  MoveL 742 to (62.2, -35.66, 5.28) mm, rotated rx 90 ry -59.82 rz 90 deg; joints [18.012, -65.128, 129.561, -160.179, 65.77, 111.765]
  MoveL 743 to (62.59, -36.33, 5.7) mm, rotated rx 90 ry -55.77 rz 90 deg; joints [17.262, -66.589, 129.722, -160.795, 64.433, 115.685]
  MoveL 744 to (62.99, -36.97, 6.17) mm, rotated rx 90 ry -51.71 rz 90 deg; joints [16.443, -67.973, 129.873, -161.501, 63.144, 119.692]
  MoveL 745 to (63.38, -37.58, 6.68) mm, rotated rx 90 ry -47.66 rz 90 deg; joints [15.557, -69.273, 130.015, -162.302, 61.911, 123.796]
  MoveL 746 to (63.82, -38.19, 7.29) mm, rotated rx 90 ry -43.28 rz 90 deg; joints [14.528, -70.576, 130.159, -163.275, 60.653, 128.346]
  MoveL 747 to (64.25, -38.76, 7.94) mm, rotated rx 90 ry -38.89 rz 90 deg; joints [13.429, -71.764, 130.295, -164.361, 59.485, 133.017]
  MoveL 748 to (64.69, -39.27, 8.63) mm, rotated rx 90 ry -34.51 rz 90 deg; joints [12.267, -72.829, 130.424, -165.558, 58.421, 137.808]
  MoveL 749 to (65.12, -39.73, 9.35) mm, rotated rx 90 ry -30.13 rz 90 deg; joints [11.047, -73.766, 130.549, -166.865, 57.475, 142.721]
  MoveL 750 to (65.56, -40.15, 10.14) mm, rotated rx 90 ry -25.6 rz 90 deg; joints [9.732, -74.593, 130.674, -168.322, 56.634, 147.917]
  MoveL 751 to (66, -40.5, 10.96) mm, rotated rx 90 ry -21.07 rz 90 deg; joints [8.373, -75.268, 130.796, -169.878, 55.946, 153.223]
  MoveL 752 to (66.44, -40.78, 11.8) mm, rotated rx 90 ry -16.54 rz 90 deg; joints [6.977, -75.787, 130.915, -171.517, 55.423, 158.623]
  MoveL 753 to (66.88, -41, 12.66) mm, rotated rx 90 ry -12.01 rz 90 deg; joints [5.554, -76.145, 131.032, -173.221, 55.076, 164.098]
  MoveL 754 to (67.32, -41.15, 13.54) mm, rotated rx 90 ry -7.48 rz 90 deg; joints [4.115, -76.339, 131.148, -174.969, 54.913, 169.623]
  MoveL 755 to (67.76, -41.23, 14.42) mm, rotated rx 90 ry -2.95 rz 90 deg; joints [2.671, -76.366, 131.26, -176.737, 54.937, 175.174]
  MoveL 756 to (68.16, -41.25, 15.26) mm, rotated rx 90 ry 0 rz 90 deg; joints [1.719, -76.288, 131.323, -177.903, 55.053, 178.798]
  MoveL 757 to (68.57, -41.25, 16.1) mm, rotated rx 90 ry 0 rz 90 deg; joints [1.676, -76.267, 131.295, -177.955, 55.045, 178.828]
  MoveL 758 to (68.97, -41.25, 16.94) mm, rotated rx 90 ry 0 rz 90 deg; joints [1.634, -76.246, 131.266, -178.007, 55.037, 178.857]
  MoveL 759 to (69.37, -41.25, 17.77) mm, rotated rx 90 ry 0 rz 90 deg; joints [1.591, -76.225, 131.238, -178.058, 55.028, 178.887]
  MoveL 760 to (69.78, -41.25, 18.61) mm, rotated rx 90 ry 0 rz 90 deg; joints [1.548, -76.204, 131.209, -178.11, 55.02, 178.916]
  MoveL 761 to (70.18, -41.25, 19.45) mm, rotated rx 90 ry 0 rz 90 deg; joints [1.506, -76.182, 131.181, -178.162, 55.012, 178.946]
  MoveL 762 to (72.7, -41.25, 24.26) mm, rotated rx 90 ry 0 rz 90 deg; joints [1.262, -76.049, 131.001, -178.459, 54.962, 179.115]
  MoveL 763 to (75.1, -41.25, 27.7) mm, rotated rx 90 ry 0 rz 90 deg; joints [1.087, -75.919, 130.826, -178.671, 54.914, 179.236]
  MoveL 764 to (78.13, -41.25, 30.71) mm, rotated rx 90 ry 0 rz 90 deg; joints [0.934, -75.754, 130.602, -178.857, 54.854, 179.342]
  MoveL 765 to (81.19, -41.25, 33.72) mm, rotated rx 90 ry 0 rz 90 deg; joints [0.782, -75.586, 130.375, -179.042, 54.793, 179.448]
  MoveL 766 to (82.71, -41.25, 36.56) mm, rotated rx 90 ry 0 rz 90 deg; joints [0.64, -75.504, 130.263, -179.216, 54.762, 179.548]
  MoveL 767 to (83.13, -41.25, 40.01) mm, rotated rx 90 ry 0 rz 90 deg; joints [0.469, -75.482, 130.234, -179.426, 54.753, 179.669]
  MoveL 768 to (82.53, -41.25, 43.6) mm, rotated rx 90 ry 0 rz 90 deg; joints [0.291, -75.517, 130.281, -179.644, 54.765, 179.795]
  MoveL 769 to (82.18, -41.25, 44.44) mm, rotated rx 90 ry 0 rz 90 deg; joints [0.25, -75.537, 130.308, -179.694, 54.772, 179.824]
  MoveL 770 to (81.83, -41.25, 45.27) mm, rotated rx 90 ry 1.37 rz 90 deg; joints [-0.208, -75.494, 130.36, 179.746, 54.866, -178.482]
  MoveL 771 to (81.47, -41.2, 46.1) mm, rotated rx 90 ry 5.62 rz 90 deg; joints [-1.527, -75.226, 130.461, 178.141, 55.25, -173.325]
  MoveL 772 to (80.96, -41.11, 46.79) mm, rotated rx 90 ry 9.15 rz 90 deg; joints [-2.612, -74.904, 130.558, 176.838, 55.695, -169.062]
  MoveL 773 to (80.45, -40.98, 47.47) mm, rotated rx 90 ry 12.69 rz 90 deg; joints [-3.676, -74.483, 130.651, 175.577, 56.246, -164.844]
  MoveL 774 to (79.95, -40.8, 48.15) mm, rotated rx 90 ry 16.23 rz 90 deg; joints [-4.716, -73.965, 130.737, 174.367, 56.9, -160.682]
  MoveL 775 to (78.97, -40.58, 48.81) mm, rotated rx 90 ry 19.82 rz 90 deg; joints [-5.743, -73.366, 130.853, 173.198, 57.67, -156.527]
  MoveL 776 to (78, -40.32, 49.47) mm, rotated rx 90 ry 23.41 rz 90 deg; joints [-6.737, -72.67, 130.961, 172.095, 58.534, -152.445]
  MoveL 777 to (77.24, -40.22, 49.7) mm, rotated rx 90 ry 24.7 rz 90 deg; joints [-7.087, -72.418, 131.028, 171.713, 58.876, -150.995]
  MoveL 778 to (76.48, -40.11, 49.93) mm, rotated rx 90 ry 25.99 rz 90 deg; joints [-7.433, -72.154, 131.094, 171.34, 59.229, -149.556]
  MoveL 779 to (75.72, -40, 50.16) mm, rotated rx 90 ry 27.28 rz 90 deg; joints [-7.774, -71.878, 131.159, 170.977, 59.593, -148.127]
  MoveL 780 to (74.77, -39.93, 50.28) mm, rotated rx 90 ry 27.99 rz 90 deg; joints [-7.964, -71.747, 131.234, 170.777, 59.813, -147.34]
  MoveL 781 to (73.82, -39.87, 50.4) mm, rotated rx 90 ry 28.71 rz 90 deg; joints [-8.153, -71.611, 131.309, 170.579, 60.036, -146.557]
  MoveL 782 to (72.87, -39.8, 50.53) mm, rotated rx 90 ry 29.42 rz 90 deg; joints [-8.34, -71.472, 131.384, 170.384, 60.262, -145.776]
  MoveL 783 to (71.92, -39.73, 50.65) mm, rotated rx 90 ry 30.13 rz 90 deg; joints [-8.525, -71.329, 131.457, 170.192, 60.491, -144.999]
  MoveL 784 to (70.97, -39.66, 50.77) mm, rotated rx 90 ry 30.85 rz 90 deg; joints [-8.709, -71.182, 131.531, 170.003, 60.724, -144.226]
  MoveL 785 to (70.02, -39.59, 50.89) mm, rotated rx 90 ry 31.56 rz 90 deg; joints [-8.892, -71.032, 131.604, 169.817, 60.96, -143.456]
  MoveL 786 to (69.07, -39.51, 51.01) mm, rotated rx 90 ry 32.27 rz 90 deg; joints [-9.073, -70.877, 131.676, 169.633, 61.199, -142.688]
  MoveL 787 to (68.12, -39.44, 51.12) mm, rotated rx 90 ry 32.99 rz 90 deg; joints [-9.252, -70.719, 131.748, 169.452, 61.441, -141.924]
  MoveL 788 to (67.17, -39.36, 51.24) mm, rotated rx 90 ry 33.7 rz 90 deg; joints [-9.43, -70.557, 131.819, 169.274, 61.686, -141.163]
  MoveL 789 to (66.22, -39.32, 51.3) mm, rotated rx 90 ry 34.04 rz 90 deg; joints [-9.518, -70.503, 131.891, 169.187, 61.817, -140.804]
  MoveL 790 to (65.27, -39.28, 51.35) mm, rotated rx 90 ry 34.38 rz 90 deg; joints [-9.606, -70.449, 131.962, 169.101, 61.949, -140.445]
  MoveL 791 to (64.32, -39.25, 51.41) mm, rotated rx 90 ry 34.72 rz 90 deg; joints [-9.693, -70.393, 132.034, 169.015, 62.081, -140.087]
  MoveL 792 to (63.37, -39.21, 51.46) mm, rotated rx 90 ry 35.06 rz 90 deg; joints [-9.78, -70.337, 132.105, 168.93, 62.215, -139.73]
  MoveL 793 to (62.41, -39.17, 51.52) mm, rotated rx 90 ry 35.4 rz 90 deg; joints [-9.866, -70.279, 132.176, 168.846, 62.348, -139.375]
  MoveL 794 to (61.46, -39.13, 51.57) mm, rotated rx 90 ry 35.74 rz 90 deg; joints [-9.953, -70.221, 132.247, 168.762, 62.483, -139.019]
  MoveL 795 to (60.51, -39.09, 51.62) mm, rotated rx 90 ry 36.08 rz 90 deg; joints [-10.039, -70.162, 132.318, 168.679, 62.619, -138.664]
  MoveL 796 to (59.55, -39.05, 51.68) mm, rotated rx 90 ry 36.41 rz 90 deg; joints [-10.124, -70.101, 132.388, 168.596, 62.755, -138.31]
  MoveL 797 to (58.6, -39.01, 51.73) mm, rotated rx 90 ry 36.75 rz 90 deg; joints [-10.21, -70.04, 132.459, 168.514, 62.892, -137.957]
  MoveL 798 to (57.65, -39.01, 51.73) mm, rotated rx 90 ry 36.77 rz 90 deg; joints [-10.223, -70.079, 132.531, 168.503, 62.925, -137.938]
  MoveL 799 to (56.69, -39.01, 51.74) mm, rotated rx 90 ry 36.79 rz 90 deg; joints [-10.236, -70.119, 132.603, 168.491, 62.958, -137.917]
  MoveL 800 to (55.73, -39.01, 51.74) mm, rotated rx 90 ry 36.81 rz 90 deg; joints [-10.249, -70.158, 132.674, 168.48, 62.991, -137.898]
  MoveL 801 to (54.78, -39, 51.74) mm, rotated rx 90 ry 36.83 rz 90 deg; joints [-10.262, -70.198, 132.746, 168.469, 63.024, -137.878]
  MoveL 802 to (53.82, -39, 51.75) mm, rotated rx 90 ry 36.85 rz 90 deg; joints [-10.275, -70.237, 132.818, 168.457, 63.057, -137.859]
  MoveL 803 to (52.87, -39, 51.75) mm, rotated rx 90 ry 36.87 rz 90 deg; joints [-10.288, -70.276, 132.89, 168.446, 63.09, -137.84]
  MoveL 804 to (51.91, -39, 51.75) mm, rotated rx 90 ry 36.9 rz 90 deg; joints [-10.302, -70.316, 132.962, 168.435, 63.123, -137.819]
  MoveL 805 to (50.96, -38.99, 51.76) mm, rotated rx 90 ry 36.91 rz 90 deg; joints [-10.315, -70.355, 133.033, 168.423, 63.156, -137.8]
  MoveL 806 to (50, -38.99, 51.76) mm, rotated rx 90 ry 36.94 rz 90 deg; joints [-10.328, -70.394, 133.105, 168.412, 63.189, -137.781]
  MoveL 807 to (50, -39.55, 50.95) mm, rotated rx 90 ry 31.94 rz 90 deg; joints [-9.143, -71.919, 133.112, 169.592, 61.592, -143.063]
  MoveL 808 to (50, -40.03, 50.1) mm, rotated rx 90 ry 26.95 rz 90 deg; joints [-7.863, -73.276, 133.093, 170.923, 60.129, -148.499]
  MoveL 809 to (50, -40.43, 49.21) mm, rotated rx 90 ry 21.96 rz 90 deg; joints [-6.498, -74.456, 133.053, 172.398, 58.821, -154.088]
  MoveL 810 to (50, -40.76, 48.28) mm, rotated rx 90 ry 16.97 rz 90 deg; joints [-5.059, -75.448, 132.995, 174.011, 57.688, -159.823]
  MoveL 811 to (50, -41.01, 47.33) mm, rotated rx 90 ry 11.98 rz 90 deg; joints [-3.556, -76.246, 132.923, 175.747, 56.75, -165.689]
  MoveL 812 to (50, -41.17, 46.37) mm, rotated rx 90 ry 6.98 rz 90 deg; joints [-2.003, -76.843, 132.841, 177.585, 56.022, -171.665]
  MoveL 813 to (50, -41.24, 45.39) mm, rotated rx 90 ry 1.99 rz 90 deg; joints [-0.413, -77.235, 132.752, 179.499, 55.517, -177.724]
  MoveL 814 to (50, -41.25, 44.41) mm, rotated rx 90 ry 0 rz 90 deg; joints [0.258, -77.334, 132.714, -179.686, 55.381, 179.822]
  MoveL 815 to (45.62, -41.25, 43.91) mm, rotated rx 90 ry 0 rz 90 deg; joints [0.285, -77.581, 133.039, -179.654, 55.459, 179.804]
  MoveL 816 to (41.42, -41.25, 43.16) mm, rotated rx 90 ry 0 rz 90 deg; joints [0.325, -77.817, 133.349, -179.606, 55.532, 179.777]
  MoveL 817 to (38.6, -41.25, 42.58) mm, rotated rx 90 ry 0 rz 90 deg; joints [0.355, -77.977, 133.557, -179.57, 55.581, 179.757]
  MoveL 818 to (35.9, -41.25, 41.66) mm, rotated rx 90 ry 0 rz 90 deg; joints [0.404, -78.13, 133.756, -179.511, 55.627, 179.724]
  MoveL 819 to (34.18, -41.25, 39.31) mm, rotated rx 90 ry 0 rz 90 deg; joints [0.526, -78.226, 133.881, -179.363, 55.657, 179.641]
  MoveL 820 to (33.35, -41.25, 35.37) mm, rotated rx 90 ry 0 rz 90 deg; joints [0.731, -78.271, 133.939, -179.115, 55.672, 179.501]
  MoveL 821 to (33.65, -41.25, 31.56) mm, rotated rx 90 ry 0 rz 90 deg; joints [0.928, -78.25, 133.913, -178.876, 55.668, 179.366]
  MoveL 822 to (34.41, -41.25, 27.86) mm, rotated rx 90 ry 0 rz 90 deg; joints [1.119, -78.203, 133.852, -178.645, 55.656, 179.235]
  MoveL 823 to (35.45, -41.25, 23.18) mm, rotated rx 90 ry 0 rz 90 deg; joints [1.36, -78.139, 133.768, -178.352, 55.64, 179.07]
  MoveL 824 to (36.64, -41.25, 18.45) mm, rotated rx 90 ry 0 rz 90 deg; joints [1.603, -78.064, 133.671, -178.057, 55.622, 178.903]
  MoveL 825 to (36.94, -41.25, 17.47) mm, rotated rx 90 ry 0 rz 90 deg; joints [1.653, -78.046, 133.647, -177.997, 55.618, 178.868]
  MoveL 826 to (37.24, -41.25, 16.5) mm, rotated rx 90 ry 0 rz 90 deg; joints [1.703, -78.027, 133.623, -177.936, 55.613, 178.834]
  MoveL 827 to (37.53, -41.25, 15.52) mm, rotated rx 90 ry 0 rz 90 deg; joints [1.753, -78.009, 133.599, -177.876, 55.608, 178.8]
  MoveL 828 to (37.83, -41.24, 14.55) mm, rotated rx 90 ry -2.31 rz 90 deg; joints [2.533, -78.043, 133.502, -176.925, 55.498, 175.947]
  MoveL 829 to (38.13, -41.16, 13.57) mm, rotated rx 90 ry -7.28 rz 90 deg; joints [4.156, -77.984, 133.319, -174.951, 55.439, 169.855]
  MoveL 830 to (38.43, -41.02, 12.72) mm, rotated rx 90 ry -11.71 rz 90 deg; joints [5.597, -77.754, 133.151, -173.21, 55.585, 164.443]
  MoveL 831 to (38.73, -40.81, 11.87) mm, rotated rx 90 ry -16.14 rz 90 deg; joints [7.021, -77.363, 132.981, -171.512, 55.912, 159.081]
  MoveL 832 to (39.03, -40.53, 11.05) mm, rotated rx 90 ry -20.57 rz 90 deg; joints [8.417, -76.813, 132.81, -169.88, 56.412, 153.793]
  MoveL 833 to (39.33, -40.2, 10.25) mm, rotated rx 90 ry -25 rz 90 deg; joints [9.777, -76.11, 132.637, -168.329, 57.076, 148.595]
  MoveL 834 to (39.63, -39.8, 9.47) mm, rotated rx 90 ry -29.43 rz 90 deg; joints [11.09, -75.258, 132.461, -166.874, 57.89, 143.505]
  MoveL 835 to (40, -39.28, 8.64) mm, rotated rx 90 ry -34.42 rz 90 deg; joints [12.506, -74.128, 132.257, -165.363, 58.971, 137.91]
  MoveL 836 to (40.37, -38.69, 7.86) mm, rotated rx 90 ry -39.41 rz 90 deg; joints [13.843, -72.827, 132.045, -163.996, 60.205, 132.475]
  MoveL 837 to (40.74, -38.04, 7.13) mm, rotated rx 90 ry -44.41 rz 90 deg; joints [15.092, -71.368, 131.825, -162.778, 61.571, 127.199]
  MoveL 838 to (41.11, -37.32, 6.46) mm, rotated rx 90 ry -49.4 rz 90 deg; joints [16.246, -69.763, 131.594, -161.709, 63.05, 122.081]
  MoveL 839 to (41.48, -36.55, 5.85) mm, rotated rx 90 ry -54.41 rz 90 deg; joints [17.302, -68.016, 131.349, -160.783, 64.628, 117.092]
  MoveL 840 to (41.84, -35.72, 5.31) mm, rotated rx 90 ry -59.43 rz 90 deg; joints [18.249, -66.15, 131.09, -159.998, 66.28, 112.244]
  MoveL 841 to (42.21, -34.85, 4.85) mm, rotated rx 90 ry -64.44 rz 90 deg; joints [19.084, -64.176, 130.813, -159.35, 67.99, 107.521]
  MoveL 842 to (42.58, -33.95, 4.47) mm, rotated rx 90 ry -69.45 rz 90 deg; joints [19.803, -62.112, 130.519, -158.83, 69.742, 102.91]
  MoveL 843 to (42.94, -33.17, 4.21) mm, rotated rx 90 ry -73.65 rz 90 deg; joints [20.313, -60.322, 130.255, -158.491, 71.229, 99.121]
  MoveL 844 to (43.3, -32.37, 4) mm, rotated rx 90 ry -77.85 rz 90 deg; joints [20.739, -58.488, 129.978, -158.233, 72.728, 95.387]
  MoveL 845 to (43.66, -31.56, 3.86) mm, rotated rx 90 ry -82.05 rz 90 deg; joints [21.079, -56.619, 129.687, -158.055, 74.232, 91.701]
  MoveL 846 to (44.02, -30.74, 3.77) mm, rotated rx 90 ry -86.25 rz 90 deg; joints [21.333, -54.723, 129.384, -157.953, 75.735, 88.05]
  MoveL 847 to (44.51, -29.87, 3.75) mm, rotated rx 0 ry -90 rz 180 deg; joints [21.484, -53.003, 129.092, -157.928, 77.072, 84.817]
  MoveL 848 to (44.99, -29, 3.75) mm, rotated rx 0 ry -90 rz 180 deg; joints [21.476, -52.928, 129.05, -157.94, 77.102, 84.831]
  MoveL 849 to (45.47, -28.14, 3.75) mm, rotated rx 0 ry -90 rz 180 deg; joints [21.467, -52.853, 129.007, -157.951, 77.132, 84.846]
  MoveL 850 to (45.95, -27.27, 3.75) mm, rotated rx 0 ry -90 rz 180 deg; joints [21.459, -52.778, 128.965, -157.963, 77.162, 84.861]
  MoveL 851 to (47.84, -24.64, 3.75) mm, rotated rx 0 ry -90 rz 180 deg; joints [21.426, -52.538, 128.807, -158.003, 77.234, 84.899]
  MoveL 852 to (48.85, -23.61, 3.75) mm, rotated rx 0 ry -90 rz 180 deg; joints [21.408, -52.437, 128.724, -158.023, 77.25, 84.91]
  MoveL 853 to (50, -22.99, 3.75) mm, rotated rx 0 ry -90 rz 180 deg; joints [21.388, -52.36, 128.634, -158.042, 77.236, 84.91]
  MoveL 854 to (51.15, -23.61, 3.75) mm, rotated rx 0 ry -90 rz 180 deg; joints [21.368, -52.37, 128.555, -158.055, 77.151, 84.88]
  MoveL 855 to (52.16, -24.64, 3.75) mm, rotated rx 0 ry -90 rz 180 deg; joints [21.351, -52.413, 128.489, -158.063, 77.049, 84.842]
  MoveL 856 to (54.05, -27.27, 3.75) mm, rotated rx 0 ry -90 rz 180 deg; joints [21.318, -52.542, 128.371, -158.075, 76.817, 84.755]
  MoveL 857 to (54.53, -28.14, 3.75) mm, rotated rx 0 ry -90 rz 180 deg; joints [21.31, -52.589, 128.343, -158.077, 76.747, 84.728]
  MoveL 858 to (55.01, -29, 3.75) mm, rotated rx 0 ry -90 rz 180 deg; joints [21.302, -52.635, 128.314, -158.079, 76.676, 84.701]
  MoveL 859 to (55.49, -29.87, 3.75) mm, rotated rx 0 ry -90 rz 180 deg; joints [21.293, -52.681, 128.285, -158.081, 76.606, 84.675]
  MoveL 860 to (55.98, -30.74, 3.77) mm, rotated rx 90 ry -86.25 rz 90 deg; joints [21.127, -54.352, 128.505, -158.116, 75.243, 87.907]
  MoveL 861 to (56.34, -31.56, 3.86) mm, rotated rx 90 ry -82.05 rz 90 deg; joints [20.863, -56.201, 128.753, -158.223, 73.729, 91.562]
  MoveL 862 to (56.7, -32.37, 4) mm, rotated rx 90 ry -77.85 rz 90 deg; joints [20.513, -58.02, 128.989, -158.407, 72.217, 95.256]
  MoveL 863 to (57.06, -33.17, 4.21) mm, rotated rx 90 ry -73.65 rz 90 deg; joints [20.08, -59.803, 129.212, -158.67, 70.712, 98.998]
  MoveL 864 to (57.42, -33.95, 4.47) mm, rotated rx 90 ry -69.45 rz 90 deg; joints [19.563, -61.538, 129.422, -159.014, 69.221, 102.798]
  MoveL 865 to (57.79, -34.85, 4.85) mm, rotated rx 90 ry -64.44 rz 90 deg; joints [18.84, -63.54, 129.66, -159.537, 67.472, 107.424]
  MoveL 866 to (58.16, -35.72, 5.31) mm, rotated rx 90 ry -59.43 rz 90 deg; joints [18.003, -65.448, 129.881, -160.188, 65.768, 112.163]
  MoveL 867 to (58.52, -36.55, 5.85) mm, rotated rx 90 ry -54.41 rz 90 deg; joints [17.056, -67.249, 130.086, -160.974, 64.123, 117.028]
  MoveL 868 to (58.89, -37.32, 6.46) mm, rotated rx 90 ry -49.4 rz 90 deg; joints [16.003, -68.928, 130.277, -161.901, 62.555, 122.035]
  MoveL 869 to (59.26, -38.04, 7.13) mm, rotated rx 90 ry -44.41 rz 90 deg; joints [14.856, -70.466, 130.453, -162.969, 61.088, 127.169]
  MoveL 870 to (59.63, -38.69, 7.86) mm, rotated rx 90 ry -39.41 rz 90 deg; joints [13.616, -71.858, 130.619, -164.183, 59.733, 132.46]
  MoveL 871 to (60, -39.28, 8.64) mm, rotated rx 90 ry -34.42 rz 90 deg; joints [12.292, -73.092, 130.777, -165.543, 58.512, 137.908]
  MoveL 872 to (60.37, -39.8, 9.47) mm, rotated rx 90 ry -29.43 rz 90 deg; joints [10.892, -74.158, 130.928, -167.045, 57.443, 143.514]
  MoveL 873 to (60.67, -40.2, 10.25) mm, rotated rx 90 ry -25 rz 90 deg; joints [9.596, -74.957, 131.059, -168.487, 56.639, 148.61]
  MoveL 874 to (60.97, -40.53, 11.05) mm, rotated rx 90 ry -20.57 rz 90 deg; joints [8.256, -75.61, 131.188, -170.023, 55.983, 153.812]
  MoveL 875 to (61.27, -40.81, 11.87) mm, rotated rx 90 ry -16.14 rz 90 deg; joints [6.883, -76.113, 131.314, -171.638, 55.488, 159.101]
  MoveL 876 to (61.57, -41.02, 12.72) mm, rotated rx 90 ry -11.71 rz 90 deg; joints [5.484, -76.46, 131.438, -173.314, 55.162, 164.462]
  MoveL 877 to (61.87, -41.16, 13.57) mm, rotated rx 90 ry -7.28 rz 90 deg; joints [4.07, -76.649, 131.561, -175.031, 55.013, 169.87]
  MoveL 878 to (62.17, -41.24, 14.55) mm, rotated rx 90 ry -2.31 rz 90 deg; joints [2.479, -76.673, 131.698, -176.976, 55.062, 175.957]
  MoveL 879 to (62.47, -41.25, 15.52) mm, rotated rx 90 ry 0 rz 90 deg; joints [1.714, -76.607, 131.749, -177.911, 55.16, 178.806]
  MoveL 880 to (62.76, -41.25, 16.5) mm, rotated rx 90 ry 0 rz 90 deg; joints [1.665, -76.592, 131.729, -177.971, 55.154, 178.841]
  MoveL 881 to (63.06, -41.25, 17.47) mm, rotated rx 90 ry 0 rz 90 deg; joints [1.615, -76.576, 131.709, -178.032, 55.148, 178.875]
  MoveL 882 to (63.36, -41.25, 18.45) mm, rotated rx 90 ry 0 rz 90 deg; joints [1.565, -76.561, 131.689, -178.092, 55.142, 178.909]
  MoveL 883 to (64.55, -41.25, 23.18) mm, rotated rx 90 ry 0 rz 90 deg; joints [1.325, -76.501, 131.609, -178.384, 55.118, 179.076]
  MoveL 884 to (65.59, -41.25, 27.86) mm, rotated rx 90 ry 0 rz 90 deg; joints [1.088, -76.449, 131.539, -178.673, 55.097, 179.241]
  MoveL 885 to (66.35, -41.25, 31.56) mm, rotated rx 90 ry 0 rz 90 deg; joints [0.901, -76.41, 131.486, -178.901, 55.081, 179.371]
  MoveL 886 to (66.65, -41.25, 35.37) mm, rotated rx 90 ry 0 rz 90 deg; joints [0.709, -76.396, 131.468, -179.135, 55.075, 179.505]
  MoveL 887 to (65.82, -41.25, 39.31) mm, rotated rx 90 ry 0 rz 90 deg; joints [0.511, -76.445, 131.533, -179.376, 55.09, 179.643]
  MoveL 888 to (64.11, -41.25, 41.66) mm, rotated rx 90 ry 0 rz 90 deg; joints [0.394, -76.542, 131.663, -179.52, 55.122, 179.726]
  MoveL 889 to (61.4, -41.25, 42.58) mm, rotated rx 90 ry 0 rz 90 deg; joints [0.348, -76.693, 131.865, -179.576, 55.172, 179.758]
  MoveL 890 to (58.58, -41.25, 43.16) mm, rotated rx 90 ry 0 rz 90 deg; joints [0.32, -76.852, 132.075, -179.611, 55.225, 179.778]
  MoveL 891 to (54.38, -41.25, 43.91) mm, rotated rx 90 ry 0 rz 90 deg; joints [0.283, -77.087, 132.388, -179.656, 55.301, 179.804]
  MoveL 892 to (50, -41.25, 44.41) mm, rotated rx 90 ry 0 rz 90 deg; joints [0.258, -77.334, 132.714, -179.686, 55.381, 179.822]
  MoveL 893 to (50, -41.25, 34.01) mm, rotated rx 90 ry 0 rz 90 deg; joints [0.789, -77.328, 132.707, -179.041, 55.382, 179.455]
  MoveL 894 to (47.54, -41.25, 33.12) mm, rotated rx 90 ry 0 rz 90 deg; joints [0.837, -77.466, 132.888, -178.984, 55.426, 179.423]
  MoveL 895 to (45.56, -41.25, 31.05) mm, rotated rx 90 ry 0 rz 90 deg; joints [0.944, -77.576, 133.033, -178.854, 55.462, 179.35]
  MoveL 896 to (44.02, -41.25, 28.52) mm, rotated rx 90 ry 0 rz 90 deg; joints [1.075, -77.661, 133.144, -178.695, 55.49, 179.261]
  MoveL 897 to (42.9, -41.25, 25.95) mm, rotated rx 90 ry 0 rz 90 deg; joints [1.209, -77.721, 133.223, -178.534, 55.511, 179.17]
  MoveL 898 to (41.78, -41.25, 20.71) mm, rotated rx 90 ry 0 rz 90 deg; joints [1.479, -77.777, 133.297, -178.205, 55.532, 178.984]
  MoveL 899 to (41.91, -41.25, 15.28) mm, rotated rx 90 ry 0 rz 90 deg; joints [1.758, -77.761, 133.275, -177.867, 55.533, 178.792]
  MoveL 900 to (42.06, -41.23, 14.35) mm, rotated rx 90 ry -3.31 rz 90 deg; joints [2.851, -77.812, 133.158, -176.535, 55.395, 174.716]
  MoveL 901 to (42.21, -41.14, 13.42) mm, rotated rx 90 ry -8.05 rz 90 deg; joints [4.394, -77.728, 132.993, -174.659, 55.381, 168.907]
  MoveL 902 to (42.36, -40.97, 12.51) mm, rotated rx 90 ry -12.79 rz 90 deg; joints [5.926, -77.458, 132.826, -172.81, 55.579, 163.133]
  MoveL 903 to (42.51, -40.73, 11.61) mm, rotated rx 90 ry -17.52 rz 90 deg; joints [7.437, -77.003, 132.657, -171.016, 55.982, 157.42]
  MoveL 904 to (42.72, -40.43, 10.78) mm, rotated rx 90 ry -22.06 rz 90 deg; joints [8.851, -76.397, 132.488, -169.373, 56.549, 152.035]
  MoveL 905 to (42.93, -40.06, 9.96) mm, rotated rx 90 ry -26.6 rz 90 deg; joints [10.225, -75.632, 132.318, -167.82, 57.282, 146.75]
  MoveL 906 to (43.13, -39.63, 9.18) mm, rotated rx 90 ry -31.13 rz 90 deg; joints [11.547, -74.714, 132.144, -166.372, 58.167, 141.581]
  MoveL 907 to (43.34, -39.14, 8.44) mm, rotated rx 90 ry -35.67 rz 90 deg; joints [12.811, -73.651, 131.965, -165.039, 59.19, 136.539]
  MoveL 908 to (43.6, -38.61, 7.76) mm, rotated rx 90 ry -40.05 rz 90 deg; joints [13.968, -72.49, 131.783, -163.865, 60.294, 131.794]
  MoveL 909 to (43.86, -38.03, 7.12) mm, rotated rx 90 ry -44.43 rz 90 deg; joints [15.057, -71.209, 131.594, -162.806, 61.497, 127.171]
  MoveL 910 to (44.12, -37.41, 6.53) mm, rotated rx 90 ry -48.81 rz 90 deg; joints [16.073, -69.815, 131.397, -161.861, 62.786, 122.671]
  MoveL 911 to (44.38, -36.74, 5.99) mm, rotated rx 90 ry -53.19 rz 90 deg; joints [17.011, -68.318, 131.19, -161.029, 64.149, 118.286]
  MoveL 912 to (44.68, -36.11, 5.55) mm, rotated rx 90 ry -57.11 rz 90 deg; joints [17.78, -66.894, 130.99, -160.379, 65.418, 114.453]
  MoveL 913 to (44.99, -35.45, 5.16) mm, rotated rx 90 ry -61.03 rz 90 deg; joints [18.482, -65.401, 130.78, -159.812, 66.726, 110.702]
  MoveL 914 to (45.3, -34.76, 4.81) mm, rotated rx 90 ry -64.95 rz 90 deg; joints [19.115, -63.846, 130.559, -159.328, 68.067, 107.025]
  MoveL 915 to (45.7, -34.02, 4.49) mm, rotated rx 90 ry -69.07 rz 90 deg; joints [19.701, -62.151, 130.31, -158.905, 69.498, 103.234]
  MoveL 916 to (46.1, -33.25, 4.23) mm, rotated rx 90 ry -73.19 rz 90 deg; joints [20.208, -60.404, 130.049, -158.565, 70.948, 99.508]
  MoveL 917 to (46.5, -32.47, 4.03) mm, rotated rx 90 ry -77.31 rz 90 deg; joints [20.634, -58.615, 129.776, -158.304, 72.41, 95.837]
  MoveL 918 to (47.02, -31.63, 3.87) mm, rotated rx 90 ry -81.68 rz 90 deg; joints [20.994, -56.674, 129.464, -158.113, 73.964, 91.991]
  MoveL 919 to (47.54, -30.77, 3.78) mm, rotated rx 90 ry -86.05 rz 90 deg; joints [21.262, -54.706, 129.14, -158.005, 75.517, 88.185]
  MoveL 920 to (48.06, -29.92, 3.75) mm, rotated rx 0 ry -90 rz 180 deg; joints [21.422, -52.903, 128.832, -157.978, 76.919, 84.769]
  MoveL 921 to (49.06, -28.63, 3.75) mm, rotated rx 0 ry -90 rz 180 deg; joints [21.405, -52.783, 128.748, -157.999, 76.951, 84.787]
  MoveL 922 to (50, -27.82, 3.75) mm, rotated rx 0 ry -90 rz 180 deg; joints [21.388, -52.699, 128.673, -158.016, 76.958, 84.795]
  MoveL 923 to (50.94, -28.63, 3.75) mm, rotated rx 0 ry -90 rz 180 deg; joints [21.372, -52.729, 128.61, -158.025, 76.871, 84.763]
  MoveL 924 to (51.94, -29.92, 3.75) mm, rotated rx 0 ry -90 rz 180 deg; joints [21.355, -52.789, 128.546, -158.032, 76.754, 84.719]
  MoveL 925 to (52.46, -30.77, 3.78) mm, rotated rx 90 ry -86.05 rz 90 deg; joints [21.177, -54.553, 128.778, -158.072, 75.315, 88.126]
  MoveL 926 to (52.98, -31.63, 3.87) mm, rotated rx 90 ry -81.68 rz 90 deg; joints [20.892, -56.477, 129.025, -158.192, 73.729, 91.926]
  MoveL 927 to (53.5, -32.47, 4.03) mm, rotated rx 90 ry -77.31 rz 90 deg; joints [20.516, -58.368, 129.258, -158.395, 72.144, 95.77]
  MoveL 928 to (53.9, -33.25, 4.23) mm, rotated rx 90 ry -73.19 rz 90 deg; joints [20.079, -60.115, 129.472, -158.664, 70.663, 99.441]
  MoveL 929 to (54.3, -34.02, 4.49) mm, rotated rx 90 ry -69.07 rz 90 deg; joints [19.562, -61.816, 129.674, -159.011, 69.197, 103.17]
  MoveL 930 to (54.7, -34.76, 4.81) mm, rotated rx 90 ry -64.95 rz 90 deg; joints [18.967, -63.463, 129.863, -159.442, 67.752, 106.965]
  MoveL 931 to (55.01, -35.45, 5.16) mm, rotated rx 90 ry -61.03 rz 90 deg; joints [18.329, -64.976, 130.037, -159.93, 66.405, 110.648]
  MoveL 932 to (55.32, -36.11, 5.55) mm, rotated rx 90 ry -57.11 rz 90 deg; joints [17.623, -66.426, 130.201, -160.5, 65.092, 114.407]
  MoveL 933 to (55.62, -36.74, 5.99) mm, rotated rx 90 ry -53.19 rz 90 deg; joints [16.851, -67.806, 130.356, -161.155, 63.821, 118.247]
  MoveL 934 to (55.88, -37.41, 6.53) mm, rotated rx 90 ry -48.81 rz 90 deg; joints [15.913, -69.261, 130.525, -161.988, 62.461, 122.641]
  MoveL 935 to (56.14, -38.03, 7.12) mm, rotated rx 90 ry -44.43 rz 90 deg; joints [14.9, -70.611, 130.684, -162.932, 61.176, 127.151]
  MoveL 936 to (56.4, -38.61, 7.76) mm, rotated rx 90 ry -40.05 rz 90 deg; joints [13.816, -71.849, 130.835, -163.99, 59.978, 131.782]
  MoveL 937 to (56.66, -39.14, 8.44) mm, rotated rx 90 ry -35.67 rz 90 deg; joints [12.665, -72.966, 130.98, -165.161, 58.88, 136.536]
  MoveL 938 to (56.87, -39.63, 9.18) mm, rotated rx 90 ry -31.13 rz 90 deg; joints [11.41, -73.991, 131.127, -166.489, 57.865, 141.585]
  MoveL 939 to (57.07, -40.06, 9.96) mm, rotated rx 90 ry -26.6 rz 90 deg; joints [10.099, -74.872, 131.271, -167.93, 56.986, 146.758]
  MoveL 940 to (57.28, -40.43, 10.78) mm, rotated rx 90 ry -22.06 rz 90 deg; joints [8.739, -75.602, 131.411, -169.473, 56.26, 152.047]
  MoveL 941 to (57.49, -40.73, 11.61) mm, rotated rx 90 ry -17.52 rz 90 deg; joints [7.34, -76.175, 131.548, -171.104, 55.697, 157.434]
  MoveL 942 to (57.64, -40.97, 12.51) mm, rotated rx 90 ry -12.79 rz 90 deg; joints [5.847, -76.604, 131.695, -172.882, 55.298, 163.146]
  MoveL 943 to (57.79, -41.14, 13.42) mm, rotated rx 90 ry -8.05 rz 90 deg; joints [4.333, -76.853, 131.839, -174.714, 55.101, 168.918]
  MoveL 944 to (57.94, -41.23, 14.35) mm, rotated rx 90 ry -3.31 rz 90 deg; joints [2.811, -76.918, 131.981, -176.572, 55.111, 174.723]
  MoveL 945 to (58.09, -41.25, 15.28) mm, rotated rx 90 ry 0 rz 90 deg; joints [1.733, -76.851, 132.075, -177.89, 55.242, 178.797]
  MoveL 946 to (58.22, -41.25, 20.71) mm, rotated rx 90 ry 0 rz 90 deg; joints [1.458, -76.852, 132.076, -178.225, 55.237, 178.988]
  MoveL 947 to (57.1, -41.25, 25.95) mm, rotated rx 90 ry 0 rz 90 deg; joints [1.193, -76.922, 132.169, -178.548, 55.256, 179.172]
  MoveL 948 to (55.98, -41.25, 28.52) mm, rotated rx 90 ry 0 rz 90 deg; joints [1.064, -76.987, 132.256, -178.705, 55.275, 179.262]
  MoveL 949 to (54.44, -41.25, 31.05) mm, rotated rx 90 ry 0 rz 90 deg; joints [0.937, -77.076, 132.374, -178.86, 55.303, 179.351]
  MoveL 950 to (52.46, -41.25, 33.12) mm, rotated rx 90 ry 0 rz 90 deg; joints [0.833, -77.19, 132.524, -178.987, 55.338, 179.424]
  MoveL 951 to (50, -41.25, 34.01) mm, rotated rx 90 ry 0 rz 90 deg; joints [0.789, -77.328, 132.707, -179.041, 55.382, 179.455]
  MoveL 952 to (50, -86.25, 34.01) mm, rotated rx 90 ry 0 rz 90 deg; joints [0.789, -79.797, 131.591, -178.995, 51.799, 179.379]
  Sollgeschwindigkeit (200.0 mm/s)
  MoveL 953 to (48.17, -86.25, 38.44) mm, rotated rx 90 ry 0 rz 90 deg; joints [0.564, -79.907, 131.729, -179.282, 51.824, 179.556]
  MoveL 954 to (46.35, -86.25, 42.86) mm, rotated rx 90 ry 0 rz 90 deg; joints [0.338, -80.017, 131.865, -179.57, 51.848, 179.734]
  MoveL 955 to (44.53, -85.85, 51.72) mm, rotated rx 90 ry 6.86 rz 90 deg; joints [-2.25, -79.646, 132.15, 177.165, 52.538, -171.412]
  MoveL 956 to (42.7, -82.81, 64.37) mm, rotated rx 90 ry 20.14 rz 90 deg; joints [-6.807, -77.603, 132.547, 171.703, 55.227, -155.106]
  MoveL 957 to (40.88, -76.95, 75.98) mm, rotated rx 90 ry 33.42 rz 90 deg; joints [-10.816, -74.04, 132.838, 167.409, 59.412, -140.098]
  MoveL 958 to (39.05, -68.58, 85.93) mm, rotated rx 90 ry 46.7 rz 90 deg; joints [-14.061, -69.153, 132.929, 164.401, 64.618, -126.48]
  MoveL 959 to (37.23, -58.15, 93.7) mm, rotated rx 90 ry 59.97 rz 90 deg; joints [-16.402, -63.219, 132.732, 162.556, 70.381, -114.004]
  MoveL 960 to (35.4, -46.21, 98.86) mm, rotated rx 90 ry 73.25 rz 90 deg; joints [-17.763, -56.576, 132.191, 161.7, 76.315, -102.275]
  MoveL 961 to (33.58, -33.41, 101.15) mm, rotated rx 90 ry 86.53 rz 90 deg; joints [-18.107, -49.598, 131.303, 161.714, 82.118, -90.877]
  MoveL 962 to (31.75, -26.73, 101.25) mm, rotated rx 0 ry 90 rz 0 deg; joints [-18.048, -47.549, 131.064, 161.844, 83.835, -87.983]
  MoveL 963 to (29.93, -22.3, 101.25) mm, rotated rx 0 ry 90 rz 0 deg; joints [-18.076, -47.253, 131.124, 161.827, 84.174, -88.092]
  MoveL 964 to (28.1, -17.88, 101.25) mm, rotated rx 0 ry 90 rz 0 deg; joints [-18.104, -46.956, 131.182, 161.81, 84.513, -88.2]
  MoveL 965 to (26.28, -13.45, 101.25) mm, rotated rx 0 ry 90 rz 0 deg; joints [-18.132, -46.657, 131.238, 161.792, 84.851, -88.309]
  MoveL 966 to (24.45, -9.03, 101.25) mm, rotated rx 0 ry 90 rz 0 deg; joints [-18.16, -46.356, 131.292, 161.773, 85.188, -88.418]
  MoveL 967 to (22.63, -4.6, 101.25) mm, rotated rx 0 ry 90 rz 0 deg; joints [-18.188, -46.054, 131.343, 161.754, 85.525, -88.527]
  Sollgeschwindigkeit (50.0 mm/s)
  MoveL 968 to (22.63, -4.6, 56.25) mm, rotated rx 0 ry 90 rz 0 deg; joints [-16.036, -46.315, 132.346, 163.927, 86.186, -88.902]
  MoveL 969 to (25.24, -8.42, 56.25) mm, rotated rx 0 ry 90 rz 0 deg; joints [-16, -46.561, 132.227, 163.956, 85.834, -88.803]
  MoveL 970 to (28.39, -11.75, 56.25) mm, rotated rx 0 ry 90 rz 0 deg; joints [-15.957, -46.757, 132.057, 163.992, 85.481, -88.705]
  MoveL 971 to (31.96, -14.9, 56.25) mm, rotated rx 0 ry 90 rz 0 deg; joints [-15.908, -46.928, 131.852, 164.033, 85.119, -88.605]
  MoveL 972 to (34.49, -17.04, 56.25) mm, rotated rx 0 ry 90 rz 0 deg; joints [-15.873, -47.041, 131.704, 164.061, 84.867, -88.536]
  MoveL 973 to (37.11, -19.32, 56.25) mm, rotated rx 0 ry 90 rz 0 deg; joints [-15.838, -47.162, 131.551, 164.09, 84.603, -88.464]
  MoveL 974 to (39.78, -21.76, 56.25) mm, rotated rx 0 ry 90 rz 0 deg; joints [-15.801, -47.292, 131.396, 164.119, 84.327, -88.389]
  MoveL 975 to (42.51, -24.11, 56.25) mm, rotated rx 0 ry 90 rz 0 deg; joints [-15.765, -47.413, 131.235, 164.148, 84.055, -88.315]
  MoveL 976 to (45.72, -25.96, 56.25) mm, rotated rx 0 ry 90 rz 0 deg; joints [-15.722, -47.484, 131.029, 164.183, 83.787, -88.244]
  MoveL 977 to (50, -26.64, 56.25) mm, rotated rx 0 ry 90 rz 0 deg; joints [-15.665, -47.443, 130.724, 164.233, 83.531, -88.178]
  MoveL 978 to (54.28, -25.96, 56.25) mm, rotated rx 0 ry 90 rz 0 deg; joints [-15.608, -47.298, 130.396, 164.284, 83.353, -88.135]
  MoveL 979 to (57.49, -24.11, 56.25) mm, rotated rx 0 ry 90 rz 0 deg; joints [-15.566, -47.09, 130.128, 164.324, 83.295, -88.123]
  MoveL 980 to (60.22, -21.76, 56.25) mm, rotated rx 0 ry 90 rz 0 deg; joints [-15.53, -46.856, 129.888, 164.36, 83.288, -88.126]
  MoveL 981 to (62.89, -19.32, 56.25) mm, rotated rx 0 ry 90 rz 0 deg; joints [-15.495, -46.616, 129.65, 164.395, 83.288, -88.13]
  MoveL 982 to (65.51, -17.04, 56.25) mm, rotated rx 0 ry 90 rz 0 deg; joints [-15.461, -46.39, 129.417, 164.429, 83.281, -88.133]
  MoveL 983 to (68.04, -14.9, 56.25) mm, rotated rx 0 ry 90 rz 0 deg; joints [-15.428, -46.176, 129.192, 164.462, 83.269, -88.133]
  MoveL 984 to (71.61, -11.75, 56.25) mm, rotated rx 0 ry 90 rz 0 deg; joints [-15.383, -45.867, 128.873, 164.508, 83.258, -88.136]
  MoveL 985 to (74.76, -8.42, 56.25) mm, rotated rx 0 ry 90 rz 0 deg; joints [-15.342, -45.554, 128.581, 164.549, 83.277, -88.147]
  MoveL 986 to (77.37, -4.6, 56.25) mm, rotated rx 0 ry 90 rz 0 deg; joints [-15.309, -45.218, 128.319, 164.585, 83.347, -88.17]
  MoveL 987 to (79.31, 0, 56.25) mm, rotated rx 0 ry 90 rz 0 deg; joints [-15.284, -44.839, 128.091, 164.614, 83.492, -88.213]
  MoveL 988 to (79.31, 0, 101.25) mm, rotated rx 0 ry 90 rz 0 deg; joints [-17.348, -44.556, 127.11, 162.514, 82.895, -87.768]
  END

--- program CFLines (robot KUKA KR 30 HA) ---
  BAS (#INITMOV,0)
  BAS (#VEL_PTP,100)
  BAS (#ACC_PTP,20)
  Sollgeschwindigkeit (200.0 mm/s)
  Werkzeug setzen: TOOL 0
  Referenz erstellen.: BASE 0
  $ADVANCE = 5
  $APO.CPTP = 1.000
  $APO.CDIS = 1.000
  Sollgeschwindigkeit (1000.0 mm/s)
  Frame wechseln at (1565.36, -92.38, 870.24) mm, rotated rx -90 ry 0 rz 0 deg
  Werkzeug setzen at (355.39, 32.27, 175.35) mm
  Sollgeschwindigkeit (200.0 mm/s)
  MoveL 2 to (-44.31, -80.09, -14.44) mm, rotated rx 90 ry -30.45 rz 90 deg; joints [14.986, -80.269, 119.983, -157.269, 42.006, 132.262]
  Sollgeschwindigkeit (50.0 mm/s)
  MoveL 3 to (-44.31, -41.29, 8.36) mm, rotated rx 90 ry -30.45 rz 90 deg; joints [13.945, -79.174, 121.774, -159.855, 44.406, 134.869]
  MoveL 4 to (-43.34, -41.28, 8.34) mm, rotated rx 90 ry -30.55 rz 90 deg; joints [13.96, -79.092, 121.706, -159.84, 44.423, 134.752]
  MoveL 5 to (-42.36, -41.27, 8.32) mm, rotated rx 90 ry -30.66 rz 90 deg; joints [13.975, -79.009, 121.639, -159.824, 44.441, 134.636]
  MoveL 6 to (-41.38, -41.26, 8.3) mm, rotated rx 90 ry -30.77 rz 90 deg; joints [13.99, -78.927, 121.571, -159.808, 44.458, 134.52]
  MoveL 7 to (-40.41, -41.24, 8.28) mm, rotated rx 90 ry -30.88 rz 90 deg; joints [14.005, -78.845, 121.503, -159.793, 44.475, 134.403]
  MoveL 8 to (-39.43, -41.23, 8.26) mm, rotated rx 90 ry -30.99 rz 90 deg; joints [14.019, -78.763, 121.435, -159.777, 44.492, 134.287]
  MoveL 9 to (-38.45, -41.22, 8.23) mm, rotated rx 90 ry -31.1 rz 90 deg; joints [14.034, -78.68, 121.367, -159.762, 44.51, 134.17]
  MoveL 10 to (-37.49, -41.11, 8.06) mm, rotated rx 90 ry -32 rz 90 deg; joints [14.237, -78.418, 121.326, -159.561, 44.769, 133.176]
  MoveL 11 to (-36.53, -41, 7.88) mm, rotated rx 90 ry -32.91 rz 90 deg; joints [14.437, -78.151, 121.285, -159.367, 45.032, 132.19]
  MoveL 12 to (-35.57, -40.88, 7.71) mm, rotated rx 90 ry -33.81 rz 90 deg; joints [14.633, -77.882, 121.246, -159.18, 45.298, 131.211]
  MoveL 13 to (-34.61, -40.77, 7.54) mm, rotated rx 90 ry -34.72 rz 90 deg; joints [14.826, -77.609, 121.207, -159, 45.566, 130.239]
  MoveL 14 to (-33.65, -40.65, 7.37) mm, rotated rx 90 ry -35.62 rz 90 deg; joints [15.016, -77.333, 121.169, -158.828, 45.838, 129.275]
  MoveL 15 to (-32.69, -40.53, 7.2) mm, rotated rx 90 ry -36.53 rz 90 deg; joints [15.203, -77.054, 121.132, -158.662, 46.112, 128.318]
  MoveL 16 to (-31.8, -40.31, 6.91) mm, rotated rx 90 ry -38.11 rz 90 deg; joints [15.53, -76.603, 121.127, -158.381, 46.613, 126.661]
  MoveL 17 to (-30.9, -40.08, 6.63) mm, rotated rx 90 ry -39.69 rz 90 deg; joints [15.847, -76.142, 121.124, -158.121, 47.121, 125.026]
  MoveL 18 to (-30, -39.85, 6.36) mm, rotated rx 90 ry -41.27 rz 90 deg; joints [16.154, -75.672, 121.123, -157.88, 47.638, 123.411]
  MoveL 19 to (-29.1, -39.6, 6.09) mm, rotated rx 90 ry -42.85 rz 90 deg; joints [16.451, -75.192, 121.124, -157.659, 48.161, 121.817]
  MoveL 20 to (-28.2, -39.35, 5.83) mm, rotated rx 90 ry -44.43 rz 90 deg; joints [16.737, -74.703, 121.127, -157.457, 48.692, 120.244]
  MoveL 21 to (-27.3, -39.1, 5.58) mm, rotated rx 90 ry -46.01 rz 90 deg; joints [17.012, -74.205, 121.132, -157.274, 49.229, 118.688]
  MoveL 22 to (-26.35, -38.63, 5.15) mm, rotated rx 90 ry -48.76 rz 90 deg; joints [17.473, -73.353, 121.19, -156.991, 50.188, 116.029]
  MoveL 23 to (-25.4, -38.15, 4.75) mm, rotated rx 90 ry -51.51 rz 90 deg; joints [17.901, -72.475, 121.252, -156.759, 51.164, 113.421]
  MoveL 24 to (-24.44, -37.65, 4.37) mm, rotated rx 90 ry -54.25 rz 90 deg; joints [18.296, -71.574, 121.317, -156.575, 52.154, 110.862]
  MoveL 25 to (-23.49, -37.13, 4.01) mm, rotated rx 90 ry -57 rz 90 deg; joints [18.657, -70.65, 121.386, -156.438, 53.156, 108.347]
  MoveL 26 to (-22.54, -36.6, 3.69) mm, rotated rx 90 ry -59.74 rz 90 deg; joints [18.984, -69.705, 121.456, -156.344, 54.168, 105.873]
  MoveL 27 to (-21.71, -35.91, 3.31) mm, rotated rx 90 ry -63.19 rz 90 deg; joints [19.35, -68.512, 121.573, -156.281, 55.458, 102.823]
  MoveL 28 to (-20.88, -35.2, 2.98) mm, rotated rx 90 ry -66.63 rz 90 deg; joints [19.662, -67.292, 121.692, -156.278, 56.758, 99.824]
  MoveL 29 to (-20.05, -34.47, 2.68) mm, rotated rx 90 ry -70.08 rz 90 deg; joints [19.918, -66.048, 121.81, -156.332, 58.064, 96.871]
  MoveL 30 to (-19.22, -33.72, 2.44) mm, rotated rx 90 ry -73.52 rz 90 deg; joints [20.119, -64.783, 121.926, -156.438, 59.374, 93.956]
  MoveL 31 to (-18.39, -32.96, 2.24) mm, rotated rx 90 ry -76.96 rz 90 deg; joints [20.265, -63.501, 122.04, -156.595, 60.685, 91.072]
  MoveL 32 to (-17.57, -32.18, 2.08) mm, rotated rx 90 ry -80.4 rz 90 deg; joints [20.354, -62.209, 122.151, -156.798, 61.992, 88.215]
  MoveL 33 to (-16.74, -31.41, 1.98) mm, rotated rx 90 ry -83.84 rz 90 deg; joints [20.388, -60.907, 122.258, -157.047, 63.294, 85.379]
  MoveL 34 to (-15.92, -30.62, 1.92) mm, rotated rx 90 ry -87.28 rz 90 deg; joints [20.366, -59.601, 122.36, -157.338, 64.588, 82.557]
  MoveL 35 to (-15.1, -29.83, 1.9) mm, rotated rx 0 ry -90 rz 180 deg; joints [20.307, -58.552, 122.423, -157.6, 65.606, 80.339]
  MoveL 36 to (-14.27, -29, 1.9) mm, rotated rx 0 ry -90 rz 180 deg; joints [20.294, -58.47, 122.364, -157.618, 65.624, 80.354]
  MoveL 37 to (-12.9, -27.3, 1.9) mm, rotated rx 0 ry -90 rz 180 deg; joints [20.273, -58.315, 122.266, -157.651, 65.674, 80.388]
  MoveL 38 to (-12.11, -25.32, 1.9) mm, rotated rx 0 ry -90 rz 180 deg; joints [20.261, -58.166, 122.214, -157.68, 65.761, 80.433]
  MoveL 39 to (-12.03, -23.12, 1.9) mm, rotated rx 0 ry -90 rz 180 deg; joints [20.259, -58.033, 122.217, -157.705, 65.887, 80.49]
  MoveL 40 to (-12.95, -19.92, 1.9) mm, rotated rx 0 ry -90 rz 180 deg; joints [20.274, -57.881, 122.3, -157.729, 66.107, 80.582]
  MoveL 41 to (-14.74, -17.2, 1.9) mm, rotated rx 0 ry -90 rz 180 deg; joints [20.301, -57.791, 122.448, -157.739, 66.331, 80.668]
  MoveL 42 to (-18.88, -13.11, 1.9) mm, rotated rx 0 ry -90 rz 180 deg; joints [20.366, -57.71, 122.779, -157.738, 66.724, 80.811]
  MoveL 43 to (-23.52, -9.64, 1.9) mm, rotated rx 0 ry -90 rz 180 deg; joints [20.438, -57.683, 123.144, -157.724, 67.098, 80.942]
  MoveL 44 to (-28.63, -7.16, 1.9) mm, rotated rx 0 ry -90 rz 180 deg; joints [20.518, -57.73, 123.541, -157.693, 67.433, 81.053]
  MoveL 45 to (-33.91, -5.84, 1.9) mm, rotated rx 0 ry -90 rz 180 deg; joints [20.602, -57.854, 123.946, -157.648, 67.707, 81.134]
  MoveL 46 to (-39.38, -5.04, 1.9) mm, rotated rx 0 ry -90 rz 180 deg; joints [20.689, -58.015, 124.364, -157.594, 67.957, 81.204]
  MoveL 47 to (-44.82, -4.13, 1.9) mm, rotated rx 0 ry -90 rz 180 deg; joints [20.777, -58.168, 124.778, -157.541, 68.213, 81.277]
  MoveL 48 to (-50, -2.49, 1.9) mm, rotated rx 0 ry -90 rz 180 deg; joints [20.861, -58.263, 125.173, -157.497, 68.502, 81.367]
  MoveL 49 to (-20.13, 0, 1.9) mm, rotated rx 0 ry -90 rz 180 deg; joints [20.385, -56.968, 122.909, -157.856, 67.533, 81.16]
  MoveL 50 to (-16.81, -1.76, 1.9) mm, rotated rx 0 ry -90 rz 180 deg; joints [20.333, -56.947, 122.651, -157.874, 67.306, 81.085]
  MoveL 51 to (-13.24, -2.81, 1.9) mm, rotated rx 0 ry -90 rz 180 deg; joints [20.278, -56.872, 122.374, -157.901, 67.11, 81.025]
  MoveL 52 to (-9.55, -3.6, 1.9) mm, rotated rx 0 ry -90 rz 180 deg; joints [20.221, -56.776, 122.088, -157.932, 66.925, 80.972]
  MoveL 53 to (-5.92, -4.55, 1.9) mm, rotated rx 0 ry -90 rz 180 deg; joints [20.166, -56.692, 121.806, -157.96, 66.733, 80.914]
  MoveL 54 to (-0.49, -6.86, 1.9) mm, rotated rx 0 ry -90 rz 180 deg; joints [20.083, -56.616, 121.38, -157.992, 66.396, 80.807]
  MoveL 55 to (4.66, -9.78, 1.9) mm, rotated rx 0 ry -90 rz 180 deg; joints [20.005, -56.585, 120.973, -158.014, 66.034, 80.686]
  MoveL 56 to (13.44, -15.59, 1.9) mm, rotated rx 0 ry -90 rz 180 deg; joints [19.874, -56.574, 120.272, -158.039, 65.372, 80.461]
  MoveL 57 to (22.11, -21.53, 1.9) mm, rotated rx 0 ry -90 rz 180 deg; joints [19.746, -56.567, 119.572, -158.058, 64.709, 80.235]
  MoveL 58 to (25.01, -23.64, 1.9) mm, rotated rx 0 ry -90 rz 180 deg; joints [19.704, -56.569, 119.337, -158.062, 64.481, 80.156]
  MoveL 59 to (27.81, -25.91, 1.9) mm, rotated rx 0 ry -90 rz 180 deg; joints [19.663, -56.583, 119.108, -158.063, 64.248, 80.075]
  MoveL 60 to (30.42, -28.42, 1.9) mm, rotated rx 0 ry -90 rz 180 deg; joints [19.625, -56.618, 118.891, -158.059, 64.009, 79.989]
  MoveL 61 to (30.89, -29.18, 1.9) mm, rotated rx 0 ry -90 rz 180 deg; joints [19.618, -56.642, 118.851, -158.055, 63.949, 79.965]
  MoveL 62 to (31.35, -29.93, 1.9) mm, rotated rx 0 ry -90 rz 180 deg; joints [19.612, -56.665, 118.811, -158.05, 63.889, 79.942]
  MoveL 63 to (31.82, -30.66, 1.92) mm, rotated rx 90 ry -87.11 rz 90 deg; joints [19.652, -57.669, 118.643, -157.785, 62.81, 82.317]
  MoveL 64 to (32.28, -31.38, 1.97) mm, rotated rx 90 ry -83.95 rz 90 deg; joints [19.653, -58.763, 118.458, -157.528, 61.627, 84.93]
  MoveL 65 to (32.53, -32.21, 2.09) mm, rotated rx 90 ry -80.29 rz 90 deg; joints [19.601, -60.033, 118.263, -157.273, 60.264, 87.971]
  MoveL 66 to (32.79, -33.03, 2.25) mm, rotated rx 90 ry -76.64 rz 90 deg; joints [19.488, -61.29, 118.063, -157.069, 58.898, 91.037]
  MoveL 67 to (33.04, -33.83, 2.47) mm, rotated rx 90 ry -72.98 rz 90 deg; joints [19.315, -62.531, 117.861, -156.919, 57.532, 94.135]
  MoveL 68 to (33.3, -34.62, 2.74) mm, rotated rx 90 ry -69.32 rz 90 deg; joints [19.081, -63.751, 117.657, -156.825, 56.17, 97.272]
  MoveL 69 to (33.53, -35.4, 3.07) mm, rotated rx 90 ry -65.64 rz 90 deg; joints [18.785, -64.956, 117.453, -156.793, 54.804, 100.481]
  MoveL 70 to (33.77, -36.16, 3.44) mm, rotated rx 90 ry -61.95 rz 90 deg; joints [18.429, -66.132, 117.249, -156.826, 53.449, 103.745]
  MoveL 71 to (34, -36.89, 3.86) mm, rotated rx 90 ry -58.27 rz 90 deg; joints [18.013, -67.275, 117.048, -156.931, 52.108, 107.073]
  MoveL 72 to (34.24, -37.59, 4.32) mm, rotated rx 90 ry -54.58 rz 90 deg; joints [17.538, -68.381, 116.85, -157.112, 50.788, 110.473]
  MoveL 73 to (34.47, -38.26, 4.83) mm, rotated rx 90 ry -50.9 rz 90 deg; joints [17.007, -69.446, 116.659, -157.375, 49.491, 113.953]
  MoveL 74 to (34.79, -38.88, 5.37) mm, rotated rx 90 ry -47.3 rz 90 deg; joints [16.433, -70.438, 116.472, -157.717, 48.251, 117.435]
  MoveL 75 to (35.11, -39.47, 5.95) mm, rotated rx 90 ry -43.71 rz 90 deg; joints [15.807, -71.385, 116.294, -158.149, 47.043, 121.009]
  MoveL 76 to (35.42, -40.02, 6.56) mm, rotated rx 90 ry -40.11 rz 90 deg; joints [15.131, -72.283, 116.126, -158.676, 45.874, 124.684]
  MoveL 77 to (35.74, -40.53, 7.21) mm, rotated rx 90 ry -36.52 rz 90 deg; joints [14.407, -73.131, 115.971, -159.303, 44.749, 128.465]
  MoveL 78 to (36.05, -41, 7.88) mm, rotated rx 90 ry -32.92 rz 90 deg; joints [13.637, -73.925, 115.829, -160.037, 43.673, 132.36]
  MoveL 79 to (36.35, -41.41, 8.57) mm, rotated rx 90 ry -29.38 rz 90 deg; joints [12.837, -74.653, 115.705, -160.865, 42.671, 136.307]
  MoveL 80 to (36.65, -41.79, 9.29) mm, rotated rx 90 ry -25.84 rz 90 deg; joints [11.998, -75.323, 115.597, -161.802, 41.73, 140.371]
  MoveL 81 to (36.95, -42.12, 10.03) mm, rotated rx 90 ry -22.31 rz 90 deg; joints [11.122, -75.935, 115.507, -162.85, 40.857, 144.556]
  MoveL 82 to (37.25, -42.4, 10.78) mm, rotated rx 90 ry -18.77 rz 90 deg; joints [10.212, -76.486, 115.436, -164.009, 40.059, 148.861]
  MoveL 83 to (37.54, -42.64, 11.56) mm, rotated rx 90 ry -15.23 rz 90 deg; joints [9.273, -76.975, 115.384, -165.276, 39.344, 153.282]
  MoveL 84 to (37.73, -42.83, 12.38) mm, rotated rx 90 ry -11.56 rz 90 deg; joints [8.27, -77.422, 115.361, -166.698, 38.698, 157.989]
  MoveL 85 to (37.92, -42.98, 13.2) mm, rotated rx 90 ry -7.88 rz 90 deg; joints [7.244, -77.797, 115.362, -168.223, 38.155, 162.807]
  MoveL 86 to (38.11, -43.07, 14.04) mm, rotated rx 90 ry -4.21 rz 90 deg; joints [6.197, -78.101, 115.386, -169.838, 37.722, 167.721]
  MoveL 87 to (38.3, -43.1, 14.88) mm, rotated rx 90 ry -0.54 rz 90 deg; joints [5.136, -78.331, 115.434, -171.526, 37.406, 172.714]
  MoveL 88 to (38.49, -43.1, 15.75) mm, rotated rx 90 ry 0 rz 90 deg; joints [4.946, -78.352, 115.436, -171.833, 37.365, 173.493]
  MoveL 89 to (38.64, -43.1, 20.36) mm, rotated rx 90 ry 0 rz 90 deg; joints [4.737, -78.367, 115.454, -172.176, 37.345, 173.766]
  MoveL 90 to (37.77, -43.1, 24.95) mm, rotated rx 90 ry 0 rz 90 deg; joints [4.532, -78.444, 115.549, -172.514, 37.341, 174.036]
  MoveL 91 to (35.77, -43.1, 29.07) mm, rotated rx 90 ry 0 rz 90 deg; joints [4.353, -78.589, 115.726, -172.814, 37.355, 174.277]
  MoveL 92 to (32.58, -43.1, 32.19) mm, rotated rx 90 ry 0 rz 90 deg; joints [4.222, -78.801, 115.987, -173.037, 37.39, 174.458]
  MoveL 93 to (28.47, -43.1, 34.01) mm, rotated rx 90 ry 0 rz 90 deg; joints [4.153, -79.065, 116.309, -173.159, 37.441, 174.559]
  MoveL 94 to (24.02, -43.1, 34.65) mm, rotated rx 90 ry 0 rz 90 deg; joints [4.138, -79.346, 116.649, -173.192, 37.5, 174.59]
  MoveL 95 to (13.93, -43.1, 34.2) mm, rotated rx 90 ry 0 rz 90 deg; joints [4.192, -79.974, 117.407, -173.124, 37.633, 174.545]
  MoveL 96 to (3.86, -43.1, 33.56) mm, rotated rx 90 ry 0 rz 90 deg; joints [4.257, -80.601, 118.157, -173.038, 37.76, 174.486]
  MoveL 97 to (-6.18, -43.1, 32.79) mm, rotated rx 90 ry 0 rz 90 deg; joints [4.328, -81.228, 118.898, -172.94, 37.88, 174.417]
  MoveL 98 to (-16.19, -43.1, 31.26) mm, rotated rx 90 ry 0 rz 90 deg; joints [4.436, -81.852, 119.627, -172.782, 37.996, 174.3]
  MoveL 99 to (-22.87, -43.1, 29.88) mm, rotated rx 90 ry 0 rz 90 deg; joints [4.526, -82.267, 120.109, -172.647, 38.071, 174.199]
  MoveL 100 to (-29.47, -43.1, 28.85) mm, rotated rx 90 ry 0 rz 90 deg; joints [4.601, -82.681, 120.584, -172.538, 38.14, 174.118]
  MoveL 101 to (-36.23, -43.1, 28.33) mm, rotated rx 90 ry 0 rz 90 deg; joints [4.652, -83.107, 121.071, -172.465, 38.206, 174.066]
  MoveL 102 to (-37.52, -43.1, 28.32) mm, rotated rx 90 ry 0 rz 90 deg; joints [4.657, -83.189, 121.165, -172.458, 38.218, 174.062]
  MoveL 103 to (-38.55, -43.1, 28.85) mm, rotated rx 90 ry 0 rz 90 deg; joints [4.636, -83.257, 121.243, -172.494, 38.225, 174.091]
  MoveL 104 to (-39.31, -43.1, 29.9) mm, rotated rx 90 ry 0 rz 90 deg; joints [4.588, -83.311, 121.304, -172.572, 38.227, 174.152]
  MoveL 105 to (-40.08, -43.1, 30.93) mm, rotated rx 90 ry 0 rz 90 deg; joints [4.542, -83.366, 121.365, -172.648, 38.23, 174.213]
  MoveL 106 to (-43.45, -43.1, 34.64) mm, rotated rx 90 ry 0 rz 90 deg; joints [4.375, -83.599, 121.629, -172.921, 38.243, 174.43]
  MoveL 107 to (-50, -43.1, 42.34) mm, rotated rx 90 ry 0 rz 90 deg; joints [4.024, -84.054, 122.141, -173.493, 38.267, 174.883]
  MoveL 108 to (-50, -43.1, 43.34) mm, rotated rx 90 ry 0 rz 90 deg; joints [3.976, -84.058, 122.146, -173.572, 38.263, 174.944]
  MoveL 109 to (-50, -43.1, 44.33) mm, rotated rx 90 ry 0 rz 90 deg; joints [3.927, -84.063, 122.151, -173.65, 38.259, 175.006]
  MoveL 110 to (-50, -43.1, 45.31) mm, rotated rx 90 ry 1.38 rz 90 deg; joints [3.462, -84.125, 122.168, -174.394, 38.177, 176.967]
  MoveL 111 to (-50, -43.04, 46.27) mm, rotated rx 90 ry 5.54 rz 90 deg; joints [2.151, -84.234, 122.234, -176.509, 38.051, -177.214]
  MoveL 112 to (-50, -42.91, 47.21) mm, rotated rx 90 ry 9.7 rz 90 deg; joints [0.839, -84.237, 122.333, -178.641, 38.103, -171.374]
  MoveL 113 to (-50, -42.72, 48.14) mm, rotated rx 90 ry 13.85 rz 90 deg; joints [-0.466, -84.134, 122.464, 179.248, 38.333, -165.556]
  MoveL 114 to (-50, -42.46, 49.05) mm, rotated rx 90 ry 18.01 rz 90 deg; joints [-1.756, -83.924, 122.627, 177.192, 38.737, -159.796]
  MoveL 115 to (-50, -42.13, 49.95) mm, rotated rx 90 ry 22.17 rz 90 deg; joints [-3.023, -83.608, 122.82, 175.225, 39.31, -154.131]
  MoveL 116 to (-50, -41.74, 50.81) mm, rotated rx 90 ry 26.33 rz 90 deg; joints [-4.259, -83.187, 123.042, 173.371, 40.044, -148.586]
  MoveL 117 to (-50, -41.29, 51.65) mm, rotated rx 90 ry 30.49 rz 90 deg; joints [-5.457, -82.661, 123.289, 171.654, 40.929, -143.187]
  MoveL 118 to (-50, -40.78, 52.45) mm, rotated rx 90 ry 34.65 rz 90 deg; joints [-6.609, -82.033, 123.559, 170.087, 41.953, -137.949]
  MoveL 119 to (-50, -40.21, 53.21) mm, rotated rx 90 ry 38.8 rz 90 deg; joints [-7.71, -81.305, 123.849, 168.678, 43.105, -132.878]
  MoveL 120 to (-50, -39.59, 53.93) mm, rotated rx 90 ry 42.96 rz 90 deg; joints [-8.753, -80.479, 124.155, 167.432, 44.37, -127.982]
  MoveL 121 to (-50, -38.91, 54.6) mm, rotated rx 90 ry 47.12 rz 90 deg; joints [-9.733, -79.559, 124.475, 166.346, 45.738, -123.255]
  MoveL 122 to (-50, -38.2, 55.22) mm, rotated rx 90 ry 51.28 rz 90 deg; joints [-10.646, -78.547, 124.804, 165.416, 47.194, -118.694]
  MoveL 123 to (-50, -37.43, 55.79) mm, rotated rx 90 ry 55.44 rz 90 deg; joints [-11.487, -77.447, 125.14, 164.635, 48.729, -114.287]
  MoveL 124 to (-49.04, -37.11, 56) mm, rotated rx 90 ry 57.1 rz 90 deg; joints [-11.794, -76.928, 125.204, 164.371, 49.345, -112.568]
  MoveL 125 to (-48.09, -36.79, 56.2) mm, rotated rx 90 ry 58.77 rz 90 deg; joints [-12.088, -76.398, 125.268, 164.129, 49.97, -110.869]
  MoveL 126 to (-47.13, -36.46, 56.39) mm, rotated rx 90 ry 60.43 rz 90 deg; joints [-12.368, -75.855, 125.331, 163.908, 50.603, -109.192]
  MoveL 127 to (-46.18, -36.13, 56.58) mm, rotated rx 90 ry 62.1 rz 90 deg; joints [-12.636, -75.301, 125.394, 163.708, 51.244, -107.535]
  MoveL 128 to (-45.22, -35.79, 56.75) mm, rotated rx 90 ry 63.76 rz 90 deg; joints [-12.891, -74.737, 125.456, 163.528, 51.89, -105.897]
  MoveL 129 to (-44.27, -35.45, 56.91) mm, rotated rx 90 ry 65.43 rz 90 deg; joints [-13.133, -74.161, 125.517, 163.368, 52.544, -104.278]
  MoveL 130 to (-43.31, -35.1, 57.07) mm, rotated rx 90 ry 67.09 rz 90 deg; joints [-13.361, -73.576, 125.576, 163.227, 53.202, -102.676]
  MoveL 131 to (-42.35, -34.75, 57.21) mm, rotated rx 90 ry 68.75 rz 90 deg; joints [-13.575, -72.98, 125.634, 163.104, 53.866, -101.091]
  MoveL 132 to (-41.47, -34.53, 57.29) mm, rotated rx 90 ry 69.76 rz 90 deg; joints [-13.695, -72.599, 125.645, 163.041, 54.262, -100.139]
  MoveL 133 to (-40.58, -34.31, 57.37) mm, rotated rx 90 ry 70.77 rz 90 deg; joints [-13.81, -72.213, 125.655, 162.985, 54.661, -99.191]
  MoveL 134 to (-39.69, -34.09, 57.44) mm, rotated rx 90 ry 71.78 rz 90 deg; joints [-13.92, -71.825, 125.665, 162.934, 55.06, -98.249]
  MoveL 135 to (-38.8, -33.88, 57.51) mm, rotated rx 90 ry 72.79 rz 90 deg; joints [-14.025, -71.435, 125.673, 162.89, 55.46, -97.313]
  MoveL 136 to (-37.91, -33.66, 57.58) mm, rotated rx 90 ry 73.8 rz 90 deg; joints [-14.125, -71.041, 125.681, 162.852, 55.86, -96.381]
  MoveL 137 to (-37.02, -33.43, 57.64) mm, rotated rx 90 ry 74.8 rz 90 deg; joints [-14.219, -70.644, 125.688, 162.82, 56.262, -95.453]
  MoveL 138 to (-36.13, -33.21, 57.7) mm, rotated rx 90 ry 75.81 rz 90 deg; joints [-14.309, -70.245, 125.694, 162.793, 56.663, -94.531]
  MoveL 139 to (-35.24, -32.99, 57.76) mm, rotated rx 90 ry 76.82 rz 90 deg; joints [-14.393, -69.844, 125.698, 162.773, 57.066, -93.612]
  MoveL 140 to (-34.35, -32.76, 57.8) mm, rotated rx 90 ry 77.83 rz 90 deg; joints [-14.472, -69.44, 125.702, 162.757, 57.468, -92.697]
  MoveL 141 to (-33.44, -32.63, 57.83) mm, rotated rx 90 ry 78.43 rz 90 deg; joints [-14.512, -69.179, 125.675, 162.754, 57.698, -92.153]
  MoveL 142 to (-32.52, -32.49, 57.86) mm, rotated rx 90 ry 79.03 rz 90 deg; joints [-14.551, -68.916, 125.647, 162.753, 57.928, -91.609]
  MoveL 143 to (-31.61, -32.36, 57.88) mm, rotated rx 90 ry 79.63 rz 90 deg; joints [-14.588, -68.654, 125.619, 162.754, 58.158, -91.068]
  MoveL 144 to (-30.7, -32.22, 57.91) mm, rotated rx 90 ry 80.23 rz 90 deg; joints [-14.623, -68.391, 125.59, 162.756, 58.387, -90.526]
  MoveL 145 to (-29.79, -32.09, 57.93) mm, rotated rx 90 ry 80.83 rz 90 deg; joints [-14.655, -68.128, 125.561, 162.761, 58.616, -89.987]
  MoveL 146 to (-28.87, -31.95, 57.95) mm, rotated rx 90 ry 81.44 rz 90 deg; joints [-14.687, -67.863, 125.531, 162.767, 58.845, -89.447]
  MoveL 147 to (-27.96, -31.81, 57.97) mm, rotated rx 90 ry 82.04 rz 90 deg; joints [-14.716, -67.598, 125.501, 162.775, 59.074, -88.909]
  MoveL 148 to (-27.05, -31.68, 57.99) mm, rotated rx 90 ry 82.64 rz 90 deg; joints [-14.744, -67.333, 125.471, 162.785, 59.303, -88.373]
  MoveL 149 to (-26.13, -31.54, 58.01) mm, rotated rx 90 ry 83.24 rz 90 deg; joints [-14.769, -67.068, 125.44, 162.796, 59.531, -87.836]
  MoveL 150 to (-25.21, -31.5, 58.01) mm, rotated rx 90 ry 83.43 rz 90 deg; joints [-14.769, -66.955, 125.381, 162.806, 59.583, -87.668]
  MoveL 151 to (-24.29, -31.46, 58.02) mm, rotated rx 90 ry 83.62 rz 90 deg; joints [-14.769, -66.841, 125.323, 162.815, 59.635, -87.499]
  MoveL 152 to (-23.37, -31.41, 58.02) mm, rotated rx 90 ry 83.8 rz 90 deg; joints [-14.769, -66.728, 125.264, 162.825, 59.688, -87.33]
  MoveL 153 to (-22.45, -31.37, 58.03) mm, rotated rx 90 ry 83.99 rz 90 deg; joints [-14.768, -66.615, 125.205, 162.835, 59.739, -87.161]
  MoveL 154 to (-21.53, -31.33, 58.03) mm, rotated rx 90 ry 84.18 rz 90 deg; joints [-14.768, -66.502, 125.146, 162.845, 59.791, -86.992]
  MoveL 155 to (-20.61, -31.29, 58.04) mm, rotated rx 90 ry 84.37 rz 90 deg; joints [-14.767, -66.388, 125.087, 162.855, 59.843, -86.823]
  MoveL 156 to (-19.69, -31.24, 58.04) mm, rotated rx 90 ry 84.55 rz 90 deg; joints [-14.766, -66.275, 125.028, 162.865, 59.894, -86.655]
  MoveL 157 to (-18.77, -31.2, 58.05) mm, rotated rx 90 ry 84.74 rz 90 deg; joints [-14.765, -66.162, 124.969, 162.876, 59.945, -86.486]
  MoveL 158 to (-17.85, -31.16, 58.05) mm, rotated rx 90 ry 84.93 rz 90 deg; joints [-14.764, -66.05, 124.91, 162.886, 59.996, -86.318]
  MoveL 159 to (-16.93, -31.18, 58.05) mm, rotated rx 90 ry 84.81 rz 90 deg; joints [-14.747, -66.05, 124.831, 162.892, 59.918, -86.421]
  MoveL 160 to (-16.01, -31.21, 58.04) mm, rotated rx 90 ry 84.69 rz 90 deg; joints [-14.73, -66.051, 124.753, 162.898, 59.84, -86.524]
  MoveL 161 to (-15.09, -31.24, 58.04) mm, rotated rx 90 ry 84.57 rz 90 deg; joints [-14.713, -66.052, 124.674, 162.904, 59.762, -86.626]
  MoveL 162 to (-14.17, -31.27, 58.04) mm, rotated rx 90 ry 84.45 rz 90 deg; joints [-14.696, -66.052, 124.596, 162.91, 59.684, -86.729]
  MoveL 163 to (-13.25, -31.29, 58.04) mm, rotated rx 90 ry 84.33 rz 90 deg; joints [-14.679, -66.052, 124.517, 162.916, 59.606, -86.832]
  MoveL 164 to (-12.33, -31.32, 58.03) mm, rotated rx 90 ry 84.21 rz 90 deg; joints [-14.662, -66.053, 124.439, 162.922, 59.528, -86.935]
  MoveL 165 to (-11.41, -31.35, 58.03) mm, rotated rx 90 ry 84.09 rz 90 deg; joints [-14.645, -66.053, 124.36, 162.928, 59.45, -87.039]
  MoveL 166 to (-10.49, -31.38, 58.03) mm, rotated rx 90 ry 83.97 rz 90 deg; joints [-14.628, -66.053, 124.282, 162.934, 59.372, -87.142]
  MoveL 167 to (-9.57, -31.4, 58.02) mm, rotated rx 90 ry 83.85 rz 90 deg; joints [-14.61, -66.053, 124.203, 162.94, 59.294, -87.245]
  MoveL 168 to (-8.61, -31.47, 58.02) mm, rotated rx 90 ry 83.57 rz 90 deg; joints [-14.584, -66.107, 124.111, 162.945, 59.15, -87.488]
  MoveL 169 to (-7.65, -31.53, 58.01) mm, rotated rx 90 ry 83.3 rz 90 deg; joints [-14.557, -66.161, 124.02, 162.95, 59.007, -87.73]
  MoveL 170 to (-6.69, -31.59, 58) mm, rotated rx 90 ry 83.02 rz 90 deg; joints [-14.53, -66.215, 123.928, 162.956, 58.863, -87.972]
  MoveL 171 to (-5.73, -31.66, 58) mm, rotated rx 90 ry 82.74 rz 90 deg; joints [-14.502, -66.269, 123.836, 162.962, 58.719, -88.216]
  MoveL 172 to (-4.77, -31.72, 57.99) mm, rotated rx 90 ry 82.47 rz 90 deg; joints [-14.474, -66.322, 123.744, 162.968, 58.576, -88.459]
  MoveL 173 to (-3.81, -31.78, 57.98) mm, rotated rx 90 ry 82.19 rz 90 deg; joints [-14.446, -66.374, 123.651, 162.975, 58.434, -88.702]
  MoveL 174 to (-2.85, -31.84, 57.97) mm, rotated rx 90 ry 81.91 rz 90 deg; joints [-14.417, -66.426, 123.559, 162.982, 58.291, -88.946]
  MoveL 175 to (-1.89, -31.91, 57.96) mm, rotated rx 90 ry 81.64 rz 90 deg; joints [-14.388, -66.479, 123.467, 162.99, 58.148, -89.191]
  MoveL 176 to (-0.93, -31.96, 57.95) mm, rotated rx 90 ry 81.4 rz 90 deg; joints [-14.362, -66.517, 123.376, 162.997, 58.021, -89.403]
  MoveL 177 to (0.04, -32.01, 57.94) mm, rotated rx 90 ry 81.16 rz 90 deg; joints [-14.334, -66.555, 123.286, 163.005, 57.893, -89.616]
  MoveL 178 to (1, -32.07, 57.94) mm, rotated rx 90 ry 80.92 rz 90 deg; joints [-14.307, -66.594, 123.195, 163.014, 57.766, -89.83]
  MoveL 179 to (1.97, -32.12, 57.93) mm, rotated rx 90 ry 80.68 rz 90 deg; joints [-14.279, -66.631, 123.105, 163.022, 57.639, -90.043]
  MoveL 180 to (2.93, -32.18, 57.92) mm, rotated rx 90 ry 80.44 rz 90 deg; joints [-14.252, -66.669, 123.014, 163.031, 57.511, -90.257]
  MoveL 181 to (3.9, -32.23, 57.91) mm, rotated rx 90 ry 80.2 rz 90 deg; joints [-14.223, -66.705, 122.923, 163.04, 57.385, -90.47]
  MoveL 182 to (4.86, -32.28, 57.9) mm, rotated rx 90 ry 79.95 rz 90 deg; joints [-14.195, -66.742, 122.832, 163.049, 57.258, -90.685]
  MoveL 183 to (5.82, -32.34, 57.89) mm, rotated rx 90 ry 79.71 rz 90 deg; joints [-14.166, -66.779, 122.741, 163.059, 57.131, -90.9]
  MoveL 184 to (6.8, -32.34, 57.89) mm, rotated rx 90 ry 79.72 rz 90 deg; joints [-14.156, -66.729, 122.665, 163.066, 57.105, -90.893]
  MoveL 185 to (7.78, -32.34, 57.89) mm, rotated rx 90 ry 79.72 rz 90 deg; joints [-14.145, -66.679, 122.589, 163.074, 57.078, -90.886]
  MoveL 186 to (8.76, -32.34, 57.89) mm, rotated rx 90 ry 79.73 rz 90 deg; joints [-14.135, -66.629, 122.513, 163.081, 57.051, -90.88]
  MoveL 187 to (9.74, -32.33, 57.89) mm, rotated rx 90 ry 79.73 rz 90 deg; joints [-14.124, -66.58, 122.437, 163.089, 57.024, -90.874]
  MoveL 188 to (10.72, -32.33, 57.89) mm, rotated rx 90 ry 79.73 rz 90 deg; joints [-14.114, -66.53, 122.361, 163.096, 56.997, -90.867]
  MoveL 189 to (11.7, -32.33, 57.89) mm, rotated rx 90 ry 79.74 rz 90 deg; joints [-14.104, -66.48, 122.285, 163.103, 56.97, -90.86]
  MoveL 190 to (12.68, -32.33, 57.89) mm, rotated rx 90 ry 79.74 rz 90 deg; joints [-14.093, -66.43, 122.209, 163.111, 56.943, -90.853]
  MoveL 191 to (13.66, -32.33, 57.89) mm, rotated rx 90 ry 79.75 rz 90 deg; joints [-14.083, -66.381, 122.132, 163.118, 56.916, -90.847]
  MoveL 192 to (14.64, -32.21, 57.91) mm, rotated rx 90 ry 80.3 rz 90 deg; joints [-14.112, -66.142, 122.092, 163.121, 57.111, -90.345]
  MoveL 193 to (15.62, -32.08, 57.93) mm, rotated rx 90 ry 80.85 rz 90 deg; joints [-14.14, -65.903, 122.051, 163.125, 57.305, -89.844]
  MoveL 194 to (16.6, -31.96, 57.95) mm, rotated rx 90 ry 81.4 rz 90 deg; joints [-14.166, -65.663, 122.01, 163.131, 57.5, -89.344]
  MoveL 195 to (17.58, -31.83, 57.97) mm, rotated rx 90 ry 81.95 rz 90 deg; joints [-14.191, -65.423, 121.969, 163.138, 57.694, -88.846]
  MoveL 196 to (18.56, -31.71, 57.99) mm, rotated rx 90 ry 82.5 rz 90 deg; joints [-14.215, -65.182, 121.927, 163.147, 57.888, -88.347]
  MoveL 197 to (19.54, -31.58, 58) mm, rotated rx 90 ry 83.06 rz 90 deg; joints [-14.237, -64.942, 121.885, 163.158, 58.081, -87.851]
  MoveL 198 to (20.45, -31.27, 58.04) mm, rotated rx 90 ry 84.45 rz 90 deg; joints [-14.303, -64.405, 121.899, 163.179, 58.62, -86.599]
  MoveL 199 to (21.37, -30.95, 58.07) mm, rotated rx 90 ry 85.85 rz 90 deg; joints [-14.36, -63.864, 121.912, 163.21, 59.157, -85.353]
  MoveL 200 to (22.28, -30.63, 58.08) mm, rotated rx 90 ry 87.25 rz 90 deg; joints [-14.407, -63.321, 121.922, 163.25, 59.694, -84.111]
  MoveL 201 to (23.19, -30.31, 58.1) mm, rotated rx 90 ry 88.65 rz 90 deg; joints [-14.445, -62.775, 121.929, 163.299, 60.23, -82.875]
  MoveL 202 to (24.11, -29.99, 58.1) mm, rotated rx 0 ry 90 rz 0 deg; joints [-14.472, -62.245, 121.932, 163.355, 60.744, -81.687]
  MoveL 203 to (25.02, -29.65, 58.1) mm, rotated rx 0 ry 90 rz 0 deg; joints [-14.462, -62.185, 121.863, 163.365, 60.735, -81.69]
  MoveL 204 to (29.98, -26.41, 58.1) mm, rotated rx 0 ry 90 rz 0 deg; joints [-14.407, -61.78, 121.504, 163.434, 60.77, -81.735]
  MoveL 205 to (34.51, -22.5, 58.1) mm, rotated rx 0 ry 90 rz 0 deg; joints [-14.357, -61.359, 121.182, 163.507, 60.858, -81.795]
  MoveL 206 to (38.75, -18.49, 58.1) mm, rotated rx 0 ry 90 rz 0 deg; joints [-14.311, -60.946, 120.882, 163.577, 60.96, -81.857]
  MoveL 207 to (41.21, -16.21, 58.1) mm, rotated rx 0 ry 90 rz 0 deg; joints [-14.284, -60.71, 120.707, 163.617, 61.015, -81.892]
  MoveL 208 to (43.79, -13.93, 58.1) mm, rotated rx 0 ry 90 rz 0 deg; joints [-14.256, -60.468, 120.521, 163.657, 61.064, -81.925]
  MoveL 209 to (46.77, -11.92, 58.1) mm, rotated rx 0 ry 90 rz 0 deg; joints [-14.224, -60.224, 120.3, 163.697, 61.082, -81.95]
  MoveL 210 to (49.96, -11.35, 58.1) mm, rotated rx 0 ry 90 rz 0 deg; joints [-14.19, -60.05, 120.05, 163.724, 61.004, -81.944]
  MoveL 211 to (53.16, -11.89, 58.1) mm, rotated rx 0 ry 90 rz 0 deg; joints [-14.155, -59.937, 119.788, 163.74, 60.857, -81.916]
  MoveL 212 to (55.52, -13.35, 58.1) mm, rotated rx 0 ry 90 rz 0 deg; joints [-14.13, -59.911, 119.586, 163.741, 60.685, -81.873]
  MoveL 213 to (57.54, -15.08, 58.1) mm, rotated rx 0 ry 90 rz 0 deg; joints [-14.109, -59.914, 119.408, 163.737, 60.507, -81.827]
  MoveL 214 to (59.47, -16.83, 58.1) mm, rotated rx 0 ry 90 rz 0 deg; joints [-14.088, -59.921, 119.238, 163.731, 60.333, -81.781]
  MoveL 215 to (63.69, -20.81, 58.1) mm, rotated rx 0 ry 90 rz 0 deg; joints [-14.044, -59.945, 118.861, 163.718, 59.943, -81.677]
  MoveL 216 to (68.07, -24.81, 58.1) mm, rotated rx 0 ry 90 rz 0 deg; joints [-13.998, -59.959, 118.469, 163.704, 59.546, -81.572]
  MoveL 217 to (72.84, -28.41, 58.1) mm, rotated rx 0 ry 90 rz 0 deg; joints [-13.948, -59.931, 118.047, 163.696, 59.161, -81.472]
  MoveL 218 to (73.72, -28.84, 58.1) mm, rotated rx 0 ry 90 rz 0 deg; joints [-13.939, -59.914, 117.972, 163.696, 59.104, -81.459]
  MoveL 219 to (74.59, -29.27, 58.1) mm, rotated rx 0 ry 90 rz 0 deg; joints [-13.93, -59.896, 117.897, 163.697, 59.048, -81.445]
  MoveL 220 to (75.47, -29.7, 58.1) mm, rotated rx 0 ry 90 rz 0 deg; joints [-13.921, -59.878, 117.821, 163.698, 58.991, -81.432]
  MoveL 221 to (76.34, -30.13, 58.1) mm, rotated rx 90 ry 89.44 rz 90 deg; joints [-13.898, -60.044, 117.717, 163.678, 58.729, -81.912]
  MoveL 222 to (77.22, -30.54, 58.09) mm, rotated rx 90 ry 87.65 rz 90 deg; joints [-13.835, -60.617, 117.548, 163.623, 58.007, -83.501]
  MoveL 223 to (78.09, -30.95, 58.07) mm, rotated rx 90 ry 85.85 rz 90 deg; joints [-13.757, -61.183, 117.376, 163.583, 57.286, -85.098]
  MoveL 224 to (79.05, -31.15, 58.05) mm, rotated rx 90 ry 84.99 rz 90 deg; joints [-13.708, -61.428, 117.248, 163.571, 56.921, -85.871]
  MoveL 225 to (80.01, -31.34, 58.03) mm, rotated rx 90 ry 84.12 rz 90 deg; joints [-13.656, -61.672, 117.119, 163.564, 56.555, -86.646]
  MoveL 226 to (80.97, -31.54, 58.01) mm, rotated rx 90 ry 83.25 rz 90 deg; joints [-13.601, -61.913, 116.989, 163.56, 56.19, -87.424]
  MoveL 227 to (81.93, -31.73, 57.98) mm, rotated rx 90 ry 82.38 rz 90 deg; joints [-13.542, -62.153, 116.859, 163.559, 55.826, -88.204]
  MoveL 228 to (82.88, -31.93, 57.96) mm, rotated rx 90 ry 81.52 rz 90 deg; joints [-13.48, -62.39, 116.728, 163.562, 55.463, -88.987]
  MoveL 229 to (83.84, -32.13, 57.93) mm, rotated rx 90 ry 80.65 rz 90 deg; joints [-13.414, -62.625, 116.596, 163.569, 55.1, -89.773]
  MoveL 230 to (84.78, -32.16, 57.92) mm, rotated rx 90 ry 80.52 rz 90 deg; joints [-13.396, -62.621, 116.511, 163.575, 55.02, -89.888]
  MoveL 231 to (85.73, -32.19, 57.92) mm, rotated rx 90 ry 80.39 rz 90 deg; joints [-13.378, -62.617, 116.426, 163.58, 54.939, -90.004]
  MoveL 232 to (86.67, -32.22, 57.91) mm, rotated rx 90 ry 80.26 rz 90 deg; joints [-13.36, -62.612, 116.341, 163.586, 54.859, -90.12]
  MoveL 233 to (87.62, -32.25, 57.91) mm, rotated rx 90 ry 80.13 rz 90 deg; joints [-13.342, -62.607, 116.256, 163.592, 54.779, -90.235]
  MoveL 234 to (88.56, -32.28, 57.9) mm, rotated rx 90 ry 80 rz 90 deg; joints [-13.323, -62.603, 116.171, 163.598, 54.698, -90.35]
  MoveL 235 to (89.51, -32.3, 57.9) mm, rotated rx 90 ry 79.86 rz 90 deg; joints [-13.305, -62.598, 116.086, 163.604, 54.618, -90.466]
  MoveL 236 to (90.45, -32.33, 57.89) mm, rotated rx 90 ry 79.73 rz 90 deg; joints [-13.287, -62.593, 116, 163.611, 54.538, -90.582]
  MoveL 237 to (91.39, -32.36, 57.88) mm, rotated rx 90 ry 79.6 rz 90 deg; joints [-13.268, -62.588, 115.915, 163.617, 54.458, -90.698]
  MoveL 238 to (92.34, -32.39, 57.88) mm, rotated rx 90 ry 79.47 rz 90 deg; joints [-13.25, -62.583, 115.829, 163.623, 54.378, -90.814]
  MoveL 239 to (93.27, -32.35, 57.89) mm, rotated rx 90 ry 79.67 rz 90 deg; joints [-13.255, -62.472, 115.766, 163.626, 54.424, -90.625]
  MoveL 240 to (94.2, -32.3, 57.9) mm, rotated rx 90 ry 79.88 rz 90 deg; joints [-13.26, -62.361, 115.702, 163.629, 54.47, -90.435]
  MoveL 241 to (95.14, -32.26, 57.9) mm, rotated rx 90 ry 80.08 rz 90 deg; joints [-13.265, -62.251, 115.639, 163.633, 54.515, -90.247]
  MoveL 242 to (96.07, -32.21, 57.91) mm, rotated rx 90 ry 80.28 rz 90 deg; joints [-13.27, -62.14, 115.575, 163.637, 54.561, -90.058]
  MoveL 243 to (97, -32.17, 57.92) mm, rotated rx 90 ry 80.48 rz 90 deg; joints [-13.274, -62.03, 115.511, 163.641, 54.606, -89.87]
  MoveL 244 to (97.93, -32.12, 57.93) mm, rotated rx 90 ry 80.68 rz 90 deg; joints [-13.278, -61.919, 115.447, 163.645, 54.652, -89.681]
  MoveL 245 to (98.86, -32.07, 57.94) mm, rotated rx 90 ry 80.89 rz 90 deg; joints [-13.282, -61.809, 115.383, 163.649, 54.697, -89.492]
  MoveL 246 to (99.8, -32.03, 57.94) mm, rotated rx 90 ry 81.09 rz 90 deg; joints [-13.286, -61.699, 115.319, 163.654, 54.742, -89.304]
  MoveL 247 to (100.73, -31.98, 57.95) mm, rotated rx 90 ry 81.29 rz 90 deg; joints [-13.29, -61.588, 115.254, 163.658, 54.787, -89.116]
  MoveL 248 to (101.66, -31.92, 57.96) mm, rotated rx 90 ry 81.56 rz 90 deg; joints [-13.298, -61.456, 115.195, 163.663, 54.858, -88.864]
  MoveL 249 to (102.58, -31.86, 57.97) mm, rotated rx 90 ry 81.83 rz 90 deg; joints [-13.305, -61.323, 115.135, 163.668, 54.929, -88.613]
  MoveL 250 to (103.51, -31.8, 57.98) mm, rotated rx 90 ry 82.1 rz 90 deg; joints [-13.313, -61.191, 115.075, 163.674, 54.999, -88.363]
  MoveL 251 to (104.43, -31.74, 57.98) mm, rotated rx 90 ry 82.37 rz 90 deg; joints [-13.32, -61.059, 115.015, 163.68, 55.07, -88.112]
  MoveL 252 to (105.36, -31.68, 57.99) mm, rotated rx 90 ry 82.64 rz 90 deg; joints [-13.326, -60.927, 114.955, 163.686, 55.141, -87.861]
  MoveL 253 to (106.28, -31.61, 58) mm, rotated rx 90 ry 82.91 rz 90 deg; joints [-13.332, -60.794, 114.895, 163.693, 55.211, -87.611]
  MoveL 254 to (107.21, -31.55, 58.01) mm, rotated rx 90 ry 83.18 rz 90 deg; joints [-13.338, -60.662, 114.835, 163.7, 55.281, -87.361]
  MoveL 255 to (108.13, -31.49, 58.01) mm, rotated rx 90 ry 83.45 rz 90 deg; joints [-13.344, -60.53, 114.774, 163.707, 55.35, -87.111]
  MoveL 256 to (109.06, -31.43, 58.02) mm, rotated rx 90 ry 83.73 rz 90 deg; joints [-13.349, -60.398, 114.714, 163.715, 55.42, -86.861]
  MoveL 257 to (109.99, -31.4, 58.02) mm, rotated rx 90 ry 83.86 rz 90 deg; joints [-13.347, -60.309, 114.645, 163.721, 55.438, -86.735]
  MoveL 258 to (110.92, -31.37, 58.03) mm, rotated rx 90 ry 83.99 rz 90 deg; joints [-13.344, -60.221, 114.575, 163.728, 55.456, -86.609]
  MoveL 259 to (111.85, -31.34, 58.03) mm, rotated rx 90 ry 84.13 rz 90 deg; joints [-13.342, -60.133, 114.506, 163.734, 55.474, -86.483]
  MoveL 260 to (112.78, -31.31, 58.03) mm, rotated rx 90 ry 84.26 rz 90 deg; joints [-13.34, -60.044, 114.437, 163.74, 55.492, -86.357]
  MoveL 261 to (113.71, -31.28, 58.04) mm, rotated rx 90 ry 84.39 rz 90 deg; joints [-13.337, -59.956, 114.367, 163.747, 55.509, -86.232]
  MoveL 262 to (114.64, -31.25, 58.04) mm, rotated rx 90 ry 84.53 rz 90 deg; joints [-13.335, -59.868, 114.298, 163.754, 55.527, -86.106]
  MoveL 263 to (115.57, -31.22, 58.04) mm, rotated rx 90 ry 84.66 rz 90 deg; joints [-13.332, -59.78, 114.228, 163.76, 55.544, -85.98]
  MoveL 264 to (116.5, -31.19, 58.05) mm, rotated rx 90 ry 84.8 rz 90 deg; joints [-13.329, -59.692, 114.158, 163.767, 55.562, -85.854]
  MoveL 265 to (117.44, -31.16, 58.05) mm, rotated rx 90 ry 84.93 rz 90 deg; joints [-13.327, -59.604, 114.089, 163.774, 55.579, -85.728]
  MoveL 266 to (118.37, -31.2, 58.05) mm, rotated rx 90 ry 84.76 rz 90 deg; joints [-13.31, -59.615, 114.001, 163.775, 55.481, -85.88]
  MoveL 267 to (119.3, -31.24, 58.04) mm, rotated rx 90 ry 84.58 rz 90 deg; joints [-13.292, -59.625, 113.913, 163.777, 55.384, -86.033]
  MoveL 268 to (120.23, -31.28, 58.04) mm, rotated rx 90 ry 84.41 rz 90 deg; joints [-13.275, -59.636, 113.826, 163.779, 55.287, -86.184]
  MoveL 269 to (121.17, -31.32, 58.03) mm, rotated rx 90 ry 84.23 rz 90 deg; joints [-13.258, -59.646, 113.738, 163.78, 55.19, -86.336]
  MoveL 270 to (122.1, -31.36, 58.03) mm, rotated rx 90 ry 84.06 rz 90 deg; joints [-13.24, -59.657, 113.65, 163.782, 55.093, -86.489]
  MoveL 271 to (123.03, -31.39, 58.02) mm, rotated rx 90 ry 83.89 rz 90 deg; joints [-13.223, -59.667, 113.562, 163.784, 54.996, -86.642]
  MoveL 272 to (123.96, -31.43, 58.02) mm, rotated rx 90 ry 83.71 rz 90 deg; joints [-13.205, -59.677, 113.475, 163.786, 54.899, -86.794]
  MoveL 273 to (124.89, -31.47, 58.02) mm, rotated rx 90 ry 83.54 rz 90 deg; joints [-13.188, -59.686, 113.386, 163.789, 54.802, -86.947]
  MoveL 274 to (125.83, -31.51, 58.01) mm, rotated rx 90 ry 83.37 rz 90 deg; joints [-13.17, -59.696, 113.298, 163.791, 54.706, -87.1]
  MoveL 275 to (126.75, -31.65, 58) mm, rotated rx 90 ry 82.77 rz 90 deg; joints [-13.129, -59.839, 113.186, 163.79, 54.453, -87.637]
  MoveL 276 to (127.68, -31.78, 57.98) mm, rotated rx 90 ry 82.17 rz 90 deg; joints [-13.087, -59.981, 113.073, 163.79, 54.202, -88.174]
  MoveL 277 to (128.6, -31.92, 57.96) mm, rotated rx 90 ry 81.58 rz 90 deg; joints [-13.043, -60.122, 112.96, 163.792, 53.951, -88.714]
  MoveL 278 to (129.53, -32.05, 57.94) mm, rotated rx 90 ry 80.98 rz 90 deg; joints [-12.997, -60.262, 112.847, 163.796, 53.7, -89.255]
  MoveL 279 to (130.45, -32.19, 57.92) mm, rotated rx 90 ry 80.39 rz 90 deg; joints [-12.95, -60.4, 112.733, 163.801, 53.449, -89.798]
  MoveL 280 to (131.37, -32.32, 57.89) mm, rotated rx 90 ry 79.79 rz 90 deg; joints [-12.902, -60.538, 112.619, 163.808, 53.199, -90.342]
  MoveL 281 to (132.3, -32.46, 57.87) mm, rotated rx 90 ry 79.2 rz 90 deg; joints [-12.852, -60.675, 112.505, 163.817, 52.95, -90.887]
  MoveL 282 to (133.22, -32.59, 57.84) mm, rotated rx 90 ry 78.6 rz 90 deg; joints [-12.8, -60.81, 112.39, 163.828, 52.701, -91.433]
  MoveL 283 to (134.15, -32.72, 57.81) mm, rotated rx 90 ry 78 rz 90 deg; joints [-12.747, -60.944, 112.275, 163.841, 52.452, -91.982]
  MoveL 284 to (135.05, -32.95, 57.76) mm, rotated rx 90 ry 76.99 rz 90 deg; joints [-12.66, -61.204, 112.135, 163.864, 52.053, -92.921]
  MoveL 285 to (135.95, -33.17, 57.71) mm, rotated rx 90 ry 75.98 rz 90 deg; joints [-12.568, -61.46, 111.994, 163.892, 51.656, -93.865]
  MoveL 286 to (136.85, -33.4, 57.65) mm, rotated rx 90 ry 74.97 rz 90 deg; joints [-12.472, -61.713, 111.853, 163.925, 51.26, -94.812]
  MoveL 287 to (137.75, -33.62, 57.59) mm, rotated rx 90 ry 73.95 rz 90 deg; joints [-12.372, -61.963, 111.711, 163.965, 50.865, -95.765]
  MoveL 288 to (138.65, -33.84, 57.52) mm, rotated rx 90 ry 72.94 rz 90 deg; joints [-12.267, -62.21, 111.568, 164.01, 50.472, -96.724]
  MoveL 289 to (139.56, -34.06, 57.45) mm, rotated rx 90 ry 71.93 rz 90 deg; joints [-12.158, -62.454, 111.425, 164.061, 50.08, -97.688]
  MoveL 290 to (140.46, -34.28, 57.38) mm, rotated rx 90 ry 70.92 rz 90 deg; joints [-12.045, -62.693, 111.281, 164.118, 49.691, -98.656]
  MoveL 291 to (141.36, -34.5, 57.3) mm, rotated rx 90 ry 69.9 rz 90 deg; joints [-11.928, -62.93, 111.136, 164.181, 49.303, -99.63]
  MoveL 292 to (142.26, -34.72, 57.22) mm, rotated rx 90 ry 68.89 rz 90 deg; joints [-11.806, -63.163, 110.991, 164.25, 48.917, -100.611]
  MoveL 293 to (143.23, -35.08, 57.08) mm, rotated rx 90 ry 67.21 rz 90 deg; joints [-11.6, -63.57, 110.794, 164.376, 48.298, -102.253]
  MoveL 294 to (144.19, -35.43, 56.92) mm, rotated rx 90 ry 65.53 rz 90 deg; joints [-11.382, -63.967, 110.596, 164.52, 47.684, -103.912]
  MoveL 295 to (145.16, -35.77, 56.76) mm, rotated rx 90 ry 63.84 rz 90 deg; joints [-11.153, -64.354, 110.396, 164.683, 47.077, -105.59]
  MoveL 296 to (146.13, -36.12, 56.58) mm, rotated rx 90 ry 62.16 rz 90 deg; joints [-10.913, -64.731, 110.196, 164.865, 46.476, -107.285]
  MoveL 297 to (147.1, -36.45, 56.4) mm, rotated rx 90 ry 60.48 rz 90 deg; joints [-10.662, -65.096, 109.996, 165.066, 45.884, -108.999]
  MoveL 298 to (148.06, -36.78, 56.2) mm, rotated rx 90 ry 58.8 rz 90 deg; joints [-10.4, -65.452, 109.795, 165.287, 45.298, -110.734]
  MoveL 299 to (149.03, -37.11, 56) mm, rotated rx 90 ry 57.12 rz 90 deg; joints [-10.128, -65.795, 109.594, 165.528, 44.722, -112.488]
  MoveL 300 to (150, -37.43, 55.79) mm, rotated rx 90 ry 55.44 rz 90 deg; joints [-9.846, -66.127, 109.393, 165.79, 44.155, -114.264]
  MoveL 301 to (150, -36.65, 56.29) mm, rotated rx 90 ry 59.49 rz 90 deg; joints [-10.491, -65.178, 109.681, 165.201, 45.469, -110.013]
  MoveL 302 to (150, -35.84, 56.73) mm, rotated rx 90 ry 63.54 rz 90 deg; joints [-11.074, -64.169, 109.967, 164.73, 46.827, -105.879]
  MoveL 303 to (150, -34.99, 57.11) mm, rotated rx 90 ry 67.59 rz 90 deg; joints [-11.59, -63.104, 110.25, 164.37, 48.22, -101.849]
  MoveL 304 to (149.08, -34.78, 57.2) mm, rotated rx 90 ry 68.59 rz 90 deg; joints [-11.715, -62.882, 110.396, 164.294, 48.597, -100.876]
  MoveL 305 to (148.16, -34.57, 57.28) mm, rotated rx 90 ry 69.59 rz 90 deg; joints [-11.836, -62.657, 110.542, 164.225, 48.976, -99.908]
  MoveL 306 to (147.24, -34.36, 57.35) mm, rotated rx 90 ry 70.58 rz 90 deg; joints [-11.952, -62.429, 110.687, 164.161, 49.357, -98.947]
  MoveL 307 to (146.32, -34.14, 57.43) mm, rotated rx 90 ry 71.58 rz 90 deg; joints [-12.065, -62.197, 110.832, 164.104, 49.74, -97.99]
  MoveL 308 to (145.4, -33.92, 57.5) mm, rotated rx 90 ry 72.58 rz 90 deg; joints [-12.173, -61.962, 110.976, 164.052, 50.124, -97.039]
  MoveL 309 to (144.48, -33.7, 57.56) mm, rotated rx 90 ry 73.58 rz 90 deg; joints [-12.278, -61.724, 111.12, 164.006, 50.51, -96.092]
  MoveL 310 to (143.56, -33.48, 57.63) mm, rotated rx 90 ry 74.57 rz 90 deg; joints [-12.378, -61.482, 111.263, 163.965, 50.898, -95.152]
  MoveL 311 to (142.64, -33.26, 57.69) mm, rotated rx 90 ry 75.57 rz 90 deg; joints [-12.474, -61.237, 111.405, 163.93, 51.287, -94.216]
  MoveL 312 to (141.72, -33.04, 57.74) mm, rotated rx 90 ry 76.57 rz 90 deg; joints [-12.566, -60.99, 111.547, 163.9, 51.677, -93.284]
  MoveL 313 to (140.81, -32.82, 57.79) mm, rotated rx 90 ry 77.57 rz 90 deg; joints [-12.654, -60.739, 111.688, 163.875, 52.069, -92.357]
  MoveL 314 to (139.88, -32.58, 57.84) mm, rotated rx 90 ry 78.65 rz 90 deg; joints [-12.744, -60.458, 111.834, 163.855, 52.494, -91.351]
  MoveL 315 to (138.96, -32.33, 57.89) mm, rotated rx 90 ry 79.74 rz 90 deg; joints [-12.829, -60.174, 111.978, 163.841, 52.921, -90.352]
  MoveL 316 to (138.04, -32.09, 57.93) mm, rotated rx 90 ry 80.83 rz 90 deg; joints [-12.909, -59.887, 112.122, 163.832, 53.348, -89.356]
  MoveL 317 to (137.12, -31.84, 57.97) mm, rotated rx 90 ry 81.91 rz 90 deg; joints [-12.983, -59.597, 112.265, 163.83, 53.777, -88.366]
  MoveL 318 to (136.2, -31.6, 58) mm, rotated rx 90 ry 83 rz 90 deg; joints [-13.053, -59.304, 112.407, 163.833, 54.206, -87.38]
  MoveL 319 to (135.28, -31.35, 58.03) mm, rotated rx 90 ry 84.08 rz 90 deg; joints [-13.117, -59.008, 112.548, 163.842, 54.637, -86.398]
  MoveL 320 to (134.36, -31.1, 58.05) mm, rotated rx 90 ry 85.17 rz 90 deg; joints [-13.177, -58.709, 112.687, 163.856, 55.067, -85.42]
  MoveL 321 to (133.44, -30.86, 58.07) mm, rotated rx 90 ry 86.26 rz 90 deg; joints [-13.231, -58.407, 112.826, 163.876, 55.499, -84.444]
  MoveL 322 to (132.51, -30.61, 58.09) mm, rotated rx 90 ry 87.34 rz 90 deg; joints [-13.28, -58.103, 112.963, 163.901, 55.931, -83.474]
  MoveL 323 to (131.59, -30.36, 58.09) mm, rotated rx 90 ry 88.43 rz 90 deg; joints [-13.323, -57.797, 113.099, 163.931, 56.363, -82.507]
  MoveL 324 to (130.66, -30.18, 58.1) mm, rotated rx 90 ry 89.2 rz 90 deg; joints [-13.354, -57.589, 113.218, 163.955, 56.681, -81.82]
  MoveL 325 to (129.73, -30, 58.1) mm, rotated rx 90 ry 89.98 rz 90 deg; joints [-13.382, -57.381, 113.336, 163.981, 57, -81.135]
  MoveL 326 to (128.8, -29.82, 58.1) mm, rotated rx 0 ry 90 rz 0 deg; joints [-13.391, -57.408, 113.417, 163.98, 57.053, -81.124]
  MoveL 327 to (127.87, -29.63, 58.1) mm, rotated rx 0 ry 90 rz 0 deg; joints [-13.4, -57.443, 113.497, 163.977, 57.098, -81.134]
  MoveL 328 to (126.94, -29.45, 58.1) mm, rotated rx 0 ry 90 rz 0 deg; joints [-13.409, -57.477, 113.577, 163.975, 57.144, -81.143]
  MoveL 329 to (126, -29.26, 58.1) mm, rotated rx 0 ry 90 rz 0 deg; joints [-13.418, -57.511, 113.657, 163.973, 57.189, -81.152]
  MoveL 330 to (125.07, -29.07, 58.1) mm, rotated rx 0 ry 90 rz 0 deg; joints [-13.427, -57.545, 113.737, 163.97, 57.234, -81.162]
  MoveL 331 to (124.14, -28.89, 58.1) mm, rotated rx 0 ry 90 rz 0 deg; joints [-13.436, -57.58, 113.817, 163.968, 57.279, -81.171]
  MoveL 332 to (123.21, -28.7, 58.1) mm, rotated rx 0 ry 90 rz 0 deg; joints [-13.445, -57.614, 113.897, 163.965, 57.324, -81.18]
  MoveL 333 to (122.28, -28.52, 58.1) mm, rotated rx 0 ry 90 rz 0 deg; joints [-13.454, -57.648, 113.976, 163.963, 57.37, -81.189]
  MoveL 334 to (112.79, -28.09, 58.1) mm, rotated rx 0 ry 90 rz 0 deg; joints [-13.546, -58.068, 114.771, 163.921, 57.743, -81.254]
  MoveL 335 to (105.31, -28.35, 58.1) mm, rotated rx 0 ry 90 rz 0 deg; joints [-13.62, -58.429, 115.388, 163.879, 58.001, -81.293]
  MoveL 336 to (97.84, -28.47, 58.1) mm, rotated rx 0 ry 90 rz 0 deg; joints [-13.694, -58.781, 116.004, 163.838, 58.265, -81.333]
  MoveL 337 to (90.33, -27.86, 58.1) mm, rotated rx 0 ry 90 rz 0 deg; joints [-13.769, -59.097, 116.626, 163.803, 58.572, -81.388]
  MoveL 338 to (83.04, -26.07, 58.1) mm, rotated rx 0 ry 90 rz 0 deg; joints [-13.843, -59.34, 117.24, 163.78, 58.939, -81.464]
  MoveL 339 to (76.31, -22.82, 58.1) mm, rotated rx 0 ry 90 rz 0 deg; joints [-13.913, -59.477, 117.819, 163.775, 59.373, -81.567]
  MoveL 340 to (70.21, -18.41, 58.1) mm, rotated rx 0 ry 90 rz 0 deg; joints [-13.976, -59.52, 118.355, 163.783, 59.855, -81.69]
  MoveL 341 to (64.6, -13.63, 58.1) mm, rotated rx 0 ry 90 rz 0 deg; joints [-14.034, -59.517, 118.851, 163.796, 60.343, -81.817]
  MoveL 342 to (59.22, -8.36, 58.1) mm, rotated rx 0 ry 90 rz 0 deg; joints [-14.091, -59.472, 119.33, 163.814, 60.853, -81.953]
  MoveL 343 to (57.44, -6.4, 58.1) mm, rotated rx 0 ry 90 rz 0 deg; joints [-14.11, -59.445, 119.489, 163.821, 61.036, -82.003]
  MoveL 344 to (55.61, -4.46, 58.1) mm, rotated rx 0 ry 90 rz 0 deg; joints [-14.129, -59.42, 119.652, 163.828, 61.219, -82.052]
  MoveL 345 to (53.63, -2.79, 58.1) mm, rotated rx 0 ry 90 rz 0 deg; joints [-14.15, -59.416, 119.825, 163.831, 61.391, -82.096]
  MoveL 346 to (51.57, -1.98, 58.1) mm, rotated rx 0 ry 90 rz 0 deg; joints [-14.172, -59.462, 119.996, 163.826, 61.515, -82.124]
  MoveL 347 to (49.02, -1.89, 58.1) mm, rotated rx 0 ry 90 rz 0 deg; joints [-14.2, -59.569, 120.202, 163.81, 61.613, -82.141]
  MoveL 348 to (46.8, -2.54, 58.1) mm, rotated rx 0 ry 90 rz 0 deg; joints [-14.224, -59.704, 120.374, 163.788, 61.652, -82.14]
  MoveL 349 to (43.99, -4.87, 58.1) mm, rotated rx 0 ry 90 rz 0 deg; joints [-14.254, -59.958, 120.581, 163.747, 61.612, -82.109]
  MoveL 350 to (41.45, -7.63, 58.1) mm, rotated rx 0 ry 90 rz 0 deg; joints [-14.281, -60.224, 120.761, 163.703, 61.533, -82.067]
  MoveL 351 to (38.97, -10.24, 58.1) mm, rotated rx 0 ry 90 rz 0 deg; joints [-14.308, -60.479, 120.937, 163.661, 61.46, -82.027]
  MoveL 352 to (33.45, -15.35, 58.1) mm, rotated rx 0 ry 90 rz 0 deg; joints [-14.369, -61.011, 121.333, 163.572, 61.338, -81.95]
  MoveL 353 to (27.56, -20.16, 58.1) mm, rotated rx 0 ry 90 rz 0 deg; joints [-14.434, -61.542, 121.756, 163.481, 61.243, -81.88]
  MoveL 354 to (21.1, -24.29, 58.1) mm, rotated rx 0 ry 90 rz 0 deg; joints [-14.506, -62.064, 122.226, 163.392, 61.204, -81.824]
  MoveL 355 to (13.97, -26.98, 58.1) mm, rotated rx 0 ry 90 rz 0 deg; joints [-14.586, -62.538, 122.761, 163.311, 61.275, -81.801]
  MoveL 356 to (6.39, -28.25, 58.1) mm, rotated rx 0 ry 90 rz 0 deg; joints [-14.672, -62.952, 123.343, 163.24, 61.447, -81.809]
  MoveL 357 to (-1.27, -28.47, 58.1) mm, rotated rx 0 ry 90 rz 0 deg; joints [-14.76, -63.312, 123.938, 163.178, 61.686, -81.839]
  MoveL 358 to (-8.89, -28.2, 58.1) mm, rotated rx 0 ry 90 rz 0 deg; joints [-14.849, -63.641, 124.534, 163.119, 61.953, -81.88]
  MoveL 359 to (-19.38, -28.23, 58.1) mm, rotated rx 0 ry 90 rz 0 deg; joints [-14.973, -64.116, 125.346, 163.032, 62.293, -81.926]
  MoveL 360 to (-29.7, -29.91, 58.1) mm, rotated rx 0 ry 90 rz 0 deg; joints [-15.097, -64.68, 126.123, 162.927, 62.514, -81.932]
  MoveL 361 to (-30.62, -30.15, 58.1) mm, rotated rx 90 ry 89.33 rz 90 deg; joints [-15.09, -64.985, 126.155, 162.892, 62.252, -82.516]
  MoveL 362 to (-31.55, -30.4, 58.09) mm, rotated rx 90 ry 88.27 rz 90 deg; joints [-15.068, -65.434, 126.164, 162.848, 61.829, -83.444]
  MoveL 363 to (-32.47, -30.64, 58.08) mm, rotated rx 90 ry 87.2 rz 90 deg; joints [-15.04, -65.881, 126.172, 162.81, 61.405, -84.373]
  MoveL 364 to (-33.39, -30.88, 58.07) mm, rotated rx 90 ry 86.14 rz 90 deg; joints [-15.007, -66.328, 126.178, 162.776, 60.979, -85.306]
  MoveL 365 to (-34.32, -31.12, 58.05) mm, rotated rx 90 ry 85.08 rz 90 deg; joints [-14.967, -66.773, 126.183, 162.748, 60.553, -86.241]
  MoveL 366 to (-35.24, -31.37, 58.03) mm, rotated rx 90 ry 84.02 rz 90 deg; joints [-14.922, -67.215, 126.186, 162.725, 60.127, -87.179]
  MoveL 367 to (-36.17, -31.61, 58) mm, rotated rx 90 ry 82.95 rz 90 deg; joints [-14.871, -67.656, 126.188, 162.707, 59.699, -88.12]
  MoveL 368 to (-37.09, -31.85, 57.97) mm, rotated rx 90 ry 81.89 rz 90 deg; joints [-14.815, -68.096, 126.189, 162.695, 59.271, -89.064]
  MoveL 369 to (-38.02, -32.09, 57.93) mm, rotated rx 90 ry 80.83 rz 90 deg; joints [-14.753, -68.532, 126.188, 162.688, 58.844, -90.011]
  MoveL 370 to (-38.94, -32.33, 57.89) mm, rotated rx 90 ry 79.77 rz 90 deg; joints [-14.685, -68.967, 126.186, 162.688, 58.416, -90.963]
  MoveL 371 to (-39.86, -32.57, 57.85) mm, rotated rx 90 ry 78.7 rz 90 deg; joints [-14.611, -69.4, 126.182, 162.693, 57.987, -91.919]
  MoveL 372 to (-40.78, -32.79, 57.8) mm, rotated rx 90 ry 77.69 rz 90 deg; joints [-14.536, -69.811, 126.181, 162.703, 57.582, -92.83]
  MoveL 373 to (-41.71, -33.02, 57.75) mm, rotated rx 90 ry 76.68 rz 90 deg; joints [-14.456, -70.219, 126.179, 162.719, 57.177, -93.746]
  MoveL 374 to (-42.63, -33.24, 57.69) mm, rotated rx 90 ry 75.67 rz 90 deg; joints [-14.371, -70.625, 126.176, 162.74, 56.771, -94.666]
  MoveL 375 to (-43.55, -33.47, 57.63) mm, rotated rx 90 ry 74.66 rz 90 deg; joints [-14.28, -71.029, 126.171, 162.767, 56.367, -95.59]
  MoveL 376 to (-44.47, -33.69, 57.57) mm, rotated rx 90 ry 73.65 rz 90 deg; joints [-14.185, -71.43, 126.166, 162.8, 55.962, -96.518]
  MoveL 377 to (-45.39, -33.91, 57.5) mm, rotated rx 90 ry 72.64 rz 90 deg; joints [-14.084, -71.828, 126.16, 162.838, 55.559, -97.451]
  MoveL 378 to (-46.31, -34.13, 57.43) mm, rotated rx 90 ry 71.63 rz 90 deg; joints [-13.978, -72.223, 126.153, 162.883, 55.156, -98.389]
  MoveL 379 to (-47.24, -34.35, 57.36) mm, rotated rx 90 ry 70.62 rz 90 deg; joints [-13.867, -72.615, 126.145, 162.934, 54.755, -99.332]
  MoveL 380 to (-48.16, -34.56, 57.28) mm, rotated rx 90 ry 69.61 rz 90 deg; joints [-13.751, -73.005, 126.136, 162.991, 54.354, -100.28]
  MoveL 381 to (-49.08, -34.78, 57.2) mm, rotated rx 90 ry 68.6 rz 90 deg; joints [-13.63, -73.391, 126.127, 163.055, 53.954, -101.234]
  MoveL 382 to (-50, -34.99, 57.11) mm, rotated rx 90 ry 67.59 rz 90 deg; joints [-13.504, -73.773, 126.117, 163.125, 53.556, -102.193]
  MoveL 383 to (-50, -34.14, 57.43) mm, rotated rx 90 ry 71.59 rz 90 deg; joints [-14.015, -72.432, 126.426, 162.852, 55.224, -98.433]
  MoveL 384 to (-50, -33.26, 57.69) mm, rotated rx 90 ry 75.58 rz 90 deg; joints [-14.448, -71.034, 126.725, 162.676, 56.919, -94.757]
  MoveL 385 to (-49.01, -33.11, 57.73) mm, rotated rx 90 ry 76.25 rz 90 deg; joints [-14.502, -70.743, 126.7, 162.664, 57.181, -94.145]
  MoveL 386 to (-48.02, -32.96, 57.76) mm, rotated rx 90 ry 76.92 rz 90 deg; joints [-14.553, -70.452, 126.673, 162.655, 57.443, -93.535]
  MoveL 387 to (-47.03, -32.81, 57.8) mm, rotated rx 90 ry 77.6 rz 90 deg; joints [-14.602, -70.159, 126.647, 162.649, 57.705, -92.927]
  MoveL 388 to (-46.04, -32.66, 57.83) mm, rotated rx 90 ry 78.27 rz 90 deg; joints [-14.648, -69.866, 126.62, 162.644, 57.967, -92.32]
  MoveL 389 to (-45.05, -32.51, 57.86) mm, rotated rx 90 ry 78.94 rz 90 deg; joints [-14.692, -69.572, 126.592, 162.643, 58.228, -91.715]
  MoveL 390 to (-44.06, -32.36, 57.88) mm, rotated rx 90 ry 79.61 rz 90 deg; joints [-14.734, -69.277, 126.564, 162.643, 58.489, -91.111]
  MoveL 391 to (-43.1, -32.08, 57.93) mm, rotated rx 90 ry 80.86 rz 90 deg; joints [-14.816, -68.77, 126.576, 162.643, 58.998, -89.996]
  MoveL 392 to (-42.14, -31.8, 57.98) mm, rotated rx 90 ry 82.1 rz 90 deg; joints [-14.89, -68.261, 126.587, 162.65, 59.506, -88.886]
  MoveL 393 to (-41.19, -31.52, 58.01) mm, rotated rx 90 ry 83.35 rz 90 deg; joints [-14.956, -67.748, 126.597, 162.665, 60.014, -87.781]
  MoveL 394 to (-40.23, -31.23, 58.04) mm, rotated rx 90 ry 84.6 rz 90 deg; joints [-15.014, -67.233, 126.604, 162.688, 60.522, -86.681]
  MoveL 395 to (-39.27, -30.95, 58.07) mm, rotated rx 90 ry 85.85 rz 90 deg; joints [-15.064, -66.715, 126.609, 162.718, 61.029, -85.584]
  MoveL 396 to (-38.31, -30.66, 58.08) mm, rotated rx 90 ry 87.09 rz 90 deg; joints [-15.107, -66.195, 126.612, 162.755, 61.536, -84.491]
  MoveL 397 to (-37.36, -30.36, 58.09) mm, rotated rx 90 ry 88.45 rz 90 deg; joints [-15.145, -65.63, 126.62, 162.803, 62.088, -83.306]
  MoveL 398 to (-36.41, -30.04, 58.1) mm, rotated rx 90 ry 89.81 rz 90 deg; joints [-15.174, -65.063, 126.626, 162.859, 62.64, -82.124]
  MoveL 399 to (-35.46, -29.72, 58.1) mm, rotated rx 0 ry 90 rz 0 deg; joints [-15.167, -64.929, 126.567, 162.878, 62.71, -81.961]
  MoveL 400 to (-34.51, -29.39, 58.1) mm, rotated rx 0 ry 90 rz 0 deg; joints [-15.156, -64.867, 126.498, 162.89, 62.701, -81.964]
  MoveL 401 to (-33.55, -29.07, 58.1) mm, rotated rx 0 ry 90 rz 0 deg; joints [-15.144, -64.805, 126.428, 162.902, 62.693, -81.968]
  MoveL 402 to (-32.6, -28.74, 58.1) mm, rotated rx 0 ry 90 rz 0 deg; joints [-15.132, -64.743, 126.359, 162.914, 62.684, -81.971]
  MoveL 403 to (-26.84, -26.99, 58.1) mm, rotated rx 0 ry 90 rz 0 deg; joints [-15.063, -64.38, 125.934, 162.982, 62.615, -81.986]
  MoveL 404 to (-20.97, -25.68, 58.1) mm, rotated rx 0 ry 90 rz 0 deg; joints [-14.992, -64.039, 125.495, 163.046, 62.511, -81.99]
  MoveL 405 to (-14.99, -24.94, 58.1) mm, rotated rx 0 ry 90 rz 0 deg; joints [-14.921, -63.727, 125.04, 163.103, 62.365, -81.98]
  MoveL 406 to (-8.98, -24.62, 58.1) mm, rotated rx 0 ry 90 rz 0 deg; joints [-14.85, -63.439, 124.577, 163.156, 62.188, -81.96]
  MoveL 407 to (-1.32, -24.11, 58.1) mm, rotated rx 0 ry 90 rz 0 deg; joints [-14.761, -63.065, 123.987, 163.223, 61.968, -81.936]
  MoveL 408 to (6.25, -22.91, 58.1) mm, rotated rx 0 ry 90 rz 0 deg; joints [-14.674, -62.656, 123.407, 163.294, 61.792, -81.926]
  MoveL 409 to (13.61, -20.71, 58.1) mm, rotated rx 0 ry 90 rz 0 deg; joints [-14.59, -62.2, 122.85, 163.373, 61.684, -81.938]
  MoveL 410 to (20.47, -17.3, 58.1) mm, rotated rx 0 ry 90 rz 0 deg; joints [-14.513, -61.7, 122.342, 163.459, 61.665, -81.976]
  MoveL 411 to (26.58, -12.68, 58.1) mm, rotated rx 0 ry 90 rz 0 deg; joints [-14.445, -61.168, 121.9, 163.549, 61.743, -82.042]
  MoveL 412 to (32.08, -7.26, 58.1) mm, rotated rx 0 ry 90 rz 0 deg; joints [-14.384, -60.619, 121.51, 163.642, 61.887, -82.125]
  MoveL 413 to (37.15, -1.5, 58.1) mm, rotated rx 0 ry 90 rz 0 deg; joints [-14.328, -60.071, 121.153, 163.732, 62.062, -82.215]
  MoveL 414 to (62.85, -1.5, 58.1) mm, rotated rx 0 ry 90 rz 0 deg; joints [-14.053, -58.936, 119.092, 163.903, 61.135, -82.069]
  MoveL 415 to (67.92, -7.26, 58.1) mm, rotated rx 0 ry 90 rz 0 deg; joints [-14, -59.024, 118.636, 163.879, 60.606, -81.926]
  MoveL 416 to (73.42, -12.68, 58.1) mm, rotated rx 0 ry 90 rz 0 deg; joints [-13.942, -59.069, 118.145, 163.86, 60.082, -81.787]
  MoveL 417 to (79.53, -17.3, 58.1) mm, rotated rx 0 ry 90 rz 0 deg; joints [-13.879, -59.038, 117.608, 163.85, 59.587, -81.66]
  MoveL 418 to (86.39, -20.71, 58.1) mm, rotated rx 0 ry 90 rz 0 deg; joints [-13.809, -58.905, 117.017, 163.855, 59.137, -81.553]
  MoveL 419 to (93.75, -22.91, 58.1) mm, rotated rx 0 ry 90 rz 0 deg; joints [-13.735, -58.682, 116.393, 163.874, 58.74, -81.467]
  MoveL 420 to (101.33, -24.11, 58.1) mm, rotated rx 0 ry 90 rz 0 deg; joints [-13.659, -58.396, 115.758, 163.903, 58.394, -81.4]
  MoveL 421 to (108.98, -24.62, 58.1) mm, rotated rx 0 ry 90 rz 0 deg; joints [-13.583, -58.069, 115.12, 163.937, 58.084, -81.345]
  MoveL 422 to (114.99, -24.94, 58.1) mm, rotated rx 0 ry 90 rz 0 deg; joints [-13.524, -57.806, 114.618, 163.965, 57.845, -81.303]
  MoveL 423 to (120.97, -25.68, 58.1) mm, rotated rx 0 ry 90 rz 0 deg; joints [-13.466, -57.566, 114.113, 163.986, 57.581, -81.253]
  MoveL 424 to (126.84, -26.99, 58.1) mm, rotated rx 0 ry 90 rz 0 deg; joints [-13.41, -57.358, 113.609, 164.001, 57.288, -81.192]
  MoveL 425 to (132.6, -28.74, 58.1) mm, rotated rx 0 ry 90 rz 0 deg; joints [-13.355, -57.176, 113.108, 164.009, 56.973, -81.122]
  MoveL 426 to (133.55, -29.07, 58.1) mm, rotated rx 0 ry 90 rz 0 deg; joints [-13.346, -57.148, 113.025, 164.009, 56.919, -81.11]
  MoveL 427 to (134.5, -29.39, 58.1) mm, rotated rx 0 ry 90 rz 0 deg; joints [-13.337, -57.12, 112.942, 164.01, 56.865, -81.098]
  MoveL 428 to (135.46, -29.72, 58.1) mm, rotated rx 0 ry 90 rz 0 deg; joints [-13.328, -57.091, 112.859, 164.011, 56.811, -81.086]
  MoveL 429 to (136.41, -30.04, 58.1) mm, rotated rx 90 ry 89.81 rz 90 deg; joints [-13.314, -57.122, 112.766, 164.005, 56.69, -81.245]
  MoveL 430 to (137.36, -30.36, 58.09) mm, rotated rx 90 ry 88.45 rz 90 deg; joints [-13.269, -57.516, 112.615, 163.958, 56.159, -82.452]
  MoveL 431 to (138.31, -30.66, 58.08) mm, rotated rx 90 ry 87.09 rz 90 deg; joints [-13.216, -57.906, 112.461, 163.919, 55.628, -83.663]
  MoveL 432 to (139.27, -30.95, 58.07) mm, rotated rx 90 ry 85.85 rz 90 deg; joints [-13.16, -58.257, 112.311, 163.891, 55.138, -84.78]
  MoveL 433 to (140.23, -31.23, 58.04) mm, rotated rx 90 ry 84.6 rz 90 deg; joints [-13.096, -58.604, 112.16, 163.871, 54.649, -85.902]
  MoveL 434 to (141.19, -31.52, 58.01) mm, rotated rx 90 ry 83.35 rz 90 deg; joints [-13.025, -58.948, 112.007, 163.857, 54.16, -87.029]
  MoveL 435 to (142.14, -31.8, 57.98) mm, rotated rx 90 ry 82.1 rz 90 deg; joints [-12.948, -59.289, 111.853, 163.851, 53.672, -88.161]
  MoveL 436 to (143.1, -32.08, 57.93) mm, rotated rx 90 ry 80.86 rz 90 deg; joints [-12.864, -59.625, 111.697, 163.853, 53.185, -89.299]
  MoveL 437 to (144.06, -32.36, 57.88) mm, rotated rx 90 ry 79.61 rz 90 deg; joints [-12.774, -59.958, 111.541, 163.862, 52.699, -90.443]
  MoveL 438 to (145.05, -32.51, 57.86) mm, rotated rx 90 ry 78.94 rz 90 deg; joints [-12.718, -60.111, 111.415, 163.872, 52.421, -91.06]
  MoveL 439 to (146.04, -32.66, 57.83) mm, rotated rx 90 ry 78.27 rz 90 deg; joints [-12.66, -60.263, 111.29, 163.885, 52.145, -91.678]
  MoveL 440 to (147.03, -32.81, 57.8) mm, rotated rx 90 ry 77.6 rz 90 deg; joints [-12.6, -60.414, 111.164, 163.899, 51.869, -92.298]
  MoveL 441 to (148.02, -32.96, 57.76) mm, rotated rx 90 ry 76.92 rz 90 deg; joints [-12.539, -60.563, 111.038, 163.916, 51.593, -92.921]
  MoveL 442 to (149.01, -33.11, 57.73) mm, rotated rx 90 ry 76.25 rz 90 deg; joints [-12.475, -60.711, 110.911, 163.935, 51.318, -93.545]
  MoveL 443 to (150, -33.26, 57.69) mm, rotated rx 90 ry 75.58 rz 90 deg; joints [-12.41, -60.857, 110.784, 163.957, 51.044, -94.172]
  MoveL 444 to (150, -32.38, 57.88) mm, rotated rx 90 ry 79.52 rz 90 deg; joints [-12.714, -59.686, 111.032, 163.886, 52.461, -90.495]
  MoveL 445 to (150, -31.49, 58.02) mm, rotated rx 90 ry 83.47 rz 90 deg; joints [-12.95, -58.48, 111.268, 163.894, 53.886, -86.877]
  MoveL 446 to (149.1, -31.28, 58.04) mm, rotated rx 90 ry 84.39 rz 90 deg; joints [-13.004, -58.237, 111.397, 163.904, 54.253, -86.042]
  MoveL 447 to (148.2, -31.07, 58.06) mm, rotated rx 90 ry 85.31 rz 90 deg; joints [-13.054, -57.992, 111.526, 163.917, 54.621, -85.209]
  MoveL 448 to (147.3, -30.86, 58.07) mm, rotated rx 90 ry 86.24 rz 90 deg; joints [-13.101, -57.745, 111.654, 163.934, 54.989, -84.379]
  MoveL 449 to (146.4, -30.65, 58.08) mm, rotated rx 90 ry 87.16 rz 90 deg; joints [-13.143, -57.496, 111.781, 163.956, 55.358, -83.551]
  MoveL 450 to (145.5, -30.44, 58.09) mm, rotated rx 90 ry 88.09 rz 90 deg; joints [-13.182, -57.245, 111.907, 163.98, 55.726, -82.727]
  MoveL 451 to (144.59, -30.23, 58.1) mm, rotated rx 90 ry 89.01 rz 90 deg; joints [-13.217, -56.992, 112.033, 164.009, 56.095, -81.905]
  MoveL 452 to (143.69, -30.02, 58.1) mm, rotated rx 90 ry 89.94 rz 90 deg; joints [-13.249, -56.737, 112.157, 164.041, 56.464, -81.084]
  MoveL 453 to (142.79, -29.79, 58.1) mm, rotated rx 0 ry 90 rz 0 deg; joints [-13.258, -56.75, 112.238, 164.042, 56.532, -81.039]
  MoveL 454 to (135.77, -27.37, 58.1) mm, rotated rx 0 ry 90 rz 0 deg; joints [-13.325, -56.96, 112.855, 164.037, 56.933, -81.13]
  MoveL 455 to (128.77, -24.91, 58.1) mm, rotated rx 0 ry 90 rz 0 deg; joints [-13.391, -57.164, 113.467, 164.031, 57.336, -81.221]
  MoveL 456 to (121.65, -22.8, 58.1) mm, rotated rx 0 ry 90 rz 0 deg; joints [-13.46, -57.389, 114.083, 164.02, 57.721, -81.305]
  MoveL 457 to (114.41, -21.15, 58.1) mm, rotated rx 0 ry 90 rz 0 deg; joints [-13.53, -57.641, 114.702, 164.001, 58.085, -81.381]
  MoveL 458 to (106.67, -19.69, 58.1) mm, rotated rx 0 ry 90 rz 0 deg; joints [-13.606, -57.923, 115.357, 163.976, 58.456, -81.455]
  MoveL 459 to (98.98, -17.97, 58.1) mm, rotated rx 0 ry 90 rz 0 deg; joints [-13.682, -58.186, 116.007, 163.953, 58.839, -81.535]
  MoveL 460 to (91.53, -15.41, 58.1) mm, rotated rx 0 ry 90 rz 0 deg; joints [-13.757, -58.392, 116.643, 163.938, 59.262, -81.629]
  MoveL 461 to (84.6, -11.65, 58.1) mm, rotated rx 0 ry 90 rz 0 deg; joints [-13.828, -58.508, 117.243, 163.936, 59.737, -81.743]
  MoveL 462 to (78.37, -6.77, 58.1) mm, rotated rx 0 ry 90 rz 0 deg; joints [-13.891, -58.529, 117.791, 163.948, 60.254, -81.875]
  MoveL 463 to (72.99, -1, 58.1) mm, rotated rx 0 ry 90 rz 0 deg; joints [-13.947, -58.458, 118.274, 163.971, 60.793, -82.02]
  MoveL 464 to (27.41, -0.5, 58.1) mm, rotated rx 0 ry 90 rz 0 deg; joints [-14.436, -60.443, 121.935, 163.673, 62.471, -82.289]
  MoveL 465 to (22.06, -6.37, 58.1) mm, rotated rx 0 ry 90 rz 0 deg; joints [-14.495, -61.012, 122.312, 163.578, 62.294, -82.197]
  MoveL 466 to (15.84, -11.36, 58.1) mm, rotated rx 0 ry 90 rz 0 deg; joints [-14.565, -61.57, 122.76, 163.483, 62.198, -82.126]
  MoveL 467 to (8.89, -15.22, 58.1) mm, rotated rx 0 ry 90 rz 0 deg; joints [-14.644, -62.1, 123.272, 163.392, 62.192, -82.079]
  MoveL 468 to (1.41, -17.87, 58.1) mm, rotated rx 0 ry 90 rz 0 deg; joints [-14.73, -62.585, 123.834, 163.308, 62.277, -82.059]
  MoveL 469 to (-6.33, -19.63, 58.1) mm, rotated rx 0 ry 90 rz 0 deg; joints [-14.819, -63.032, 124.42, 163.229, 62.423, -82.057]
  MoveL 470 to (-14.13, -21.1, 58.1) mm, rotated rx 0 ry 90 rz 0 deg; joints [-14.911, -63.465, 125.012, 163.15, 62.587, -82.062]
  MoveL 471 to (-21.43, -22.75, 58.1) mm, rotated rx 0 ry 90 rz 0 deg; joints [-14.998, -63.888, 125.56, 163.072, 62.719, -82.058]
  MoveL 472 to (-28.61, -24.85, 58.1) mm, rotated rx 0 ry 90 rz 0 deg; joints [-15.084, -64.334, 126.092, 162.989, 62.813, -82.043]
  MoveL 473 to (-35.67, -27.33, 58.1) mm, rotated rx 0 ry 90 rz 0 deg; joints [-15.17, -64.798, 126.608, 162.901, 62.876, -82.016]
  MoveL 474 to (-42.74, -29.78, 58.1) mm, rotated rx 0 ry 90 rz 0 deg; joints [-15.257, -65.261, 127.124, 162.813, 62.937, -81.989]
  MoveL 475 to (-43.65, -30, 58.1) mm, rotated rx 90 ry 90 rz 90 deg; joints [-15.268, -65.317, 127.19, 162.802, 62.949, -81.991]
  MoveL 476 to (-44.55, -30.21, 58.1) mm, rotated rx 90 ry 89.06 rz 90 deg; joints [-15.253, -65.722, 127.206, 162.759, 62.575, -82.802]
  MoveL 477 to (-45.46, -30.43, 58.09) mm, rotated rx 90 ry 88.13 rz 90 deg; joints [-15.234, -66.126, 127.22, 162.72, 62.2, -83.615]
  MoveL 478 to (-46.37, -30.64, 58.08) mm, rotated rx 90 ry 87.2 rz 90 deg; joints [-15.21, -66.528, 127.233, 162.685, 61.825, -84.429]
  MoveL 479 to (-47.28, -30.85, 58.07) mm, rotated rx 90 ry 86.26 rz 90 deg; joints [-15.182, -66.93, 127.245, 162.654, 61.448, -85.245]
  MoveL 480 to (-48.19, -31.07, 58.06) mm, rotated rx 90 ry 85.33 rz 90 deg; joints [-15.149, -67.331, 127.255, 162.627, 61.071, -86.063]
  MoveL 481 to (-49.09, -31.28, 58.04) mm, rotated rx 90 ry 84.4 rz 90 deg; joints [-15.112, -67.73, 127.265, 162.604, 60.693, -86.883]
  MoveL 482 to (-50, -31.49, 58.02) mm, rotated rx 90 ry 83.47 rz 90 deg; joints [-15.07, -68.128, 127.273, 162.586, 60.315, -87.706]
  MoveL 483 to (-50, -30.73, 58.08) mm, rotated rx 90 ry 86.81 rz 90 deg; joints [-15.239, -66.846, 127.485, 162.642, 61.766, -84.778]
  MoveL 484 to (-50, -29.96, 58.1) mm, rotated rx 0 ry 90 rz 0 deg; joints [-15.347, -65.6, 127.675, 162.744, 63.152, -82.015]
  MoveL 485 to (-50, -29.16, 58.1) mm, rotated rx 0 ry 90 rz 0 deg; joints [-15.347, -65.552, 127.684, 162.753, 63.207, -82.033]
  MoveL 486 to (-45.03, -27.98, 58.1) mm, rotated rx 0 ry 90 rz 0 deg; joints [-15.285, -65.258, 127.318, 162.811, 63.13, -82.041]
  MoveL 487 to (-40.36, -26.03, 58.1) mm, rotated rx 0 ry 90 rz 0 deg; joints [-15.227, -64.931, 126.981, 162.873, 63.112, -82.066]
  MoveL 488 to (-35.76, -23.86, 58.1) mm, rotated rx 0 ry 90 rz 0 deg; joints [-15.171, -64.596, 126.651, 162.937, 63.11, -82.097]
  MoveL 489 to (-31.09, -21.86, 58.1) mm, rotated rx 0 ry 90 rz 0 deg; joints [-15.114, -64.268, 126.313, 162.998, 63.091, -82.122]
  MoveL 490 to (-26.38, -19.97, 58.1) mm, rotated rx 0 ry 90 rz 0 deg; joints [-15.057, -63.946, 125.969, 163.058, 63.062, -82.143]
  MoveL 491 to (-21.65, -18.1, 58.1) mm, rotated rx 0 ry 90 rz 0 deg; joints [-15, -63.626, 125.622, 163.118, 63.03, -82.163]
  MoveL 492 to (-14.36, -15.46, 58.1) mm, rotated rx 0 ry 90 rz 0 deg; joints [-14.914, -63.147, 125.083, 163.205, 62.96, -82.187]
  MoveL 493 to (-7.03, -12.94, 58.1) mm, rotated rx 0 ry 90 rz 0 deg; joints [-14.828, -62.674, 124.536, 163.29, 62.878, -82.207]
  MoveL 494 to (0.1, -9.83, 58.1) mm, rotated rx 0 ry 90 rz 0 deg; joints [-14.745, -62.179, 124.008, 163.377, 62.834, -82.238]
  MoveL 495 to (6.7, -5.75, 58.1) mm, rotated rx 0 ry 90 rz 0 deg; joints [-14.669, -61.652, 123.526, 163.468, 62.867, -82.291]
  MoveL 496 to (12.41, -0.5, 58.1) mm, rotated rx 0 ry 90 rz 0 deg; joints [-14.604, -61.099, 123.119, 163.562, 63, -82.371]
